# B&R Automation Studio project lab2_2
Automation Studio 4.5.2.102; technology packages: Acp10Arnc0 5.2.1

## Configuration Config1

CPU 4PP065.0571-P74, AutomationRuntime D4.52, Build 4.1.2, Vc V4.52.0, Safety 1.6

### Task classes (Cpu.sw)
```
Cyclic#1:
  ncsdcctrl <- ncsdcctrl.prg
Cyclic#2:
  Program <- Program.prg
DataObjects: Arnc0sys, Acp10sys
NcDataObjects: acp10etxen <- acp10etxen.dob, gmcipvar <- GmcIpUserConfig.gmcipvar.dob, gmcipfun <- GmcIpUserConfig.gmcipfun.dob, gmcipfub <- GmcIpUserConfig.gmcipfub.dob, gmcipubr <- GmcIpUserConfig.gmcipubr.dob, gmcipusm <- GmcIpUserConfig.gmcipusm.dob, gmcipui <- GmcIpUserConfig.gmcipui.dob, gmcipus <- GmcIpUserConfig.gmcipus.dob, gmcipuc <- GmcIpUserConfig.gmcipuc.dob, gmcipsys <- GmcIpConfig.gmcipsys.dob, gmciplbr <- GmcIpConfig.gmciplbr.dob, gmcipcbr <- GmcIpConfig.gmcipcbr.dob, gmciplsm <- GmcIpConfig.gmciplsm.dob, gmcipcsm <- GmcIpConfig.gmcipcsm.dob, gmcipcfg <- GmcIpConfig.gmcipcfg.dob, gmcipiec <- GmcIpConfig.gmcipiec.dob, gmciplog <- GmcIpConfig.gmciplog.dob, gmcipesm <- GmcIpConfig.gmcipesm.dob, gmcipmxd <- GmcIpConfig.gmcipmxd.dob, gmcipmx <- GmcIpConfig.gmcipmx.dob, gAxis01a <- gAxis01obj.gAxis01a.dob, gAxis01i <- gAxis01obj.gAxis01i.dob
Binaries: udbdef, TCData, iomap, asfw, Role, ashwac, sysconf, ashwd, User, arconfig, Arnc0map, acp10cfg, Acp10map, arnc0cfg
Libraries: Acp10man, Acp10par, NcGlobal, Acp10sdc, AsBrStr, Arnc0man, DataObj, AsArLog, sys_lib, FileIO, AsArProf, AsMem, brsystem, runtime, astime, Acp10_MC, Library, asieccon, powerlnk
```

### IoMap.iom - 4PP065_0571_P74/IoMap.iom
```iecst
VAR_CONFIG
	Cyclic#1.gAxis01_DrvIf.iLifeCnt AT %IB."X20SM1436a".LifeCnt;
	Cyclic#1.gAxis01_DrvIf.iDrvOK AT %IX."X20SM1436a".DrvOk01;
	Cyclic#1.gAxis01_DrvIf.oBoostCurrent AT %QX."X20SM1436a".BoostCurrent01;
	Cyclic#1.gAxis01_DrvIf.oStandStillCurrent AT %QX."X20SM1436a".StandstillCurrent01;
	Cyclic#1.gAxis01_DrvIf.oSetTime AT %QW."X20SM1436a".SetTime01;
	Cyclic#1.gAxis01_MotorStep0 AT %QW."X20SM1436a".Motor1Step0;
	Cyclic#1.gAxis01_DiDoIf.iLifeCntDriveEnable AT %IB."X20SM1436a".LifeCnt;
	Cyclic#1.gAxis01_DiDoIf.iLifeCntDriveReady AT %IB."X20SM1436a".LifeCnt;
	Cyclic#1.gAxis01_DiDoIf.iDriveReady AT %IX."X20SM1436a".DrvOk01;
	Cyclic#1.gAxis01_DiDoIf.oDriveEnable AT %QX."X20SM1436a".DriveEnable01;
	Cyclic#1.gAxis01_EncIf1.iLifeCnt AT %IB."X20SM1436a".LifeCnt;
	Cyclic#1.gAxis01_EncIf1.iEncOK AT %IX."X20SM1436a".EncOk01;
	Cyclic#1.gAxis01_EncIf1.iActPos AT %IW."X20SM1436a".ActPos01;
	Cyclic#1.gAxis01_EncIf1.iRefPulsePos AT %IW."X20SM1436a".RefPulsePos01;
	Cyclic#1.gAxis01_EncIf1.iRefPulseCnt AT %IB."X20SM1436a".RefPulseCnt01;
	Cyclic#1.gAxis01_EncIf1.iActTime AT %IW."X20SM1436a".ActTime01;
	::stateMachine.state AT %IW."8I64xxxxxxx.00x-1".ETAD_Input;
	::stateMachine.command AT %QW."8I64xxxxxxx.00x-1".CMDD_Output;
	::stateMachine.speed AT %QW."8I64xxxxxxx.00x-1".LFRD_Output;
	::doorSM.direction AT %IX."X20DI9371".DigitalInput01;
	::doorSM.sw1 AT %IX."X20DI9371".DigitalInput02;
	::doorSM.sw2 AT %IX."X20DI9371".DigitalInput03;
	::doorSM.sw3 AT %IX."X20DI9371".DigitalInput04;
	::doorSM.sw4 AT %IX."X20DI9371".DigitalInput05;
	::ledSM.led1 AT %QX."X20DO9322".DigitalOutput02;
	::ledSM.led2 AT %QX."X20DO9322".DigitalOutput03;
	::ledSM.led3 AT %QX."X20DO9322".DigitalOutput04;
	::ledSM.led4 AT %QX."X20DO9322".DigitalOutput05;
END_VAR
```

### Acp10cfg.ncc - 4PP065_0571_P74/Motion/Acp10cfg.ncc
```
NcConfiguration (Version=5.02.1, NcSwId=Acp10)
  ACP10CF1_typ:
    cnt_nettrc_rec_drive = 1500
    bufsize_trace_upload = 1200
    tc_nc_man_task = Cyclic #1
    glob_pv_as_ncobject = Yes
    ncsys_dl_broadcast = Yes
    ncsys_dl_acp_reset = Yes
    safemc_log_err_to_ax = Yes
    network_init:
      ncsw_init_execute = Yes
      automatic_execute = No
      node_nr_warning = Yes
      net_err_before_ncact = Yes
    nettrc:
      enter_parsecrec = Yes
      enter_ncaction = Yes
      save_ring_startidx = Yes
    cam_prof_download:
      cam_dat_dl_parallel = No
      tc_cam_dl_parallel = Task class for NC Manager task
    sdc_if[0]:
      if_name = SDC_IF1
      mc_broadcast_size = 800
      mc_broadcast_extdat = No
```

### Acp10map.ncm - 4PP065_0571_P74/Motion/Acp10map.ncm
```
NcMapping (NcSwId=Acp10)
  NcObject X20SM1436_ncAXIS1 (ModuleId=X20SM1436, ModuleAddress=SDC_IF1.ST1, Type=ncAXIS, Channel=1, AcoposSimulation=Off, Disabled=TRUE, ModuleDisabled=FALSE)
  NcObject gAxis01 (ModuleId=X20SM1436a, ModuleAddress=SDC_IF1.ST2, Type=ncAXIS, Channel=1, AcoposSimulation=Off, InitParameter=gAxis01i, AcoposParameter=gAxis01a, AdditionalData=CNC_Enabled="1" , Disabled=FALSE, ModuleDisabled=FALSE)
```

### Arnc0cfg.ncc - 4PP065_0571_P74/Motion/Arnc0cfg.ncc
```
NcConfiguration (Version=5.02.1, NcSwId=Arnc0)
  ARNC0CFG_typ:
    sampling_rate = 4000
    cnt_nettrc_rec_drive = 150
    bufsize_sys_trace = 16#00005000
    enable_mp_log = Yes
    tc_nc_man_task = Cyclic #1
    bg_load = 1
    glob_pv_as_ncobject = Yes
```

### Arnc0map.ncm - 4PP065_0571_P74/Motion/Arnc0map.ncm
```
NcMapping (NcSwId=Arnc0)
  NcObject CNC1 (Type=ncCNCSYS, Channel=1, AcoposSimulation=Off, Disabled=TRUE, ModuleDisabled=FALSE)
  NcObject CNC2 (Type=ncCNCSYS, Channel=2, AcoposSimulation=Off, Disabled=TRUE, ModuleDisabled=FALSE)
  NcObject CNC3 (Type=ncCNCSYS, Channel=3, AcoposSimulation=Off, Disabled=TRUE, ModuleDisabled=FALSE)
  NcObject CNC4 (Type=ncCNCSYS, Channel=4, AcoposSimulation=Off, Disabled=TRUE, ModuleDisabled=FALSE)
  NcObject CNC5 (Type=ncCNCSYS, Channel=5, AcoposSimulation=Off, Disabled=TRUE, ModuleDisabled=FALSE)
  NcObject CNC6 (Type=ncCNCSYS, Channel=6, AcoposSimulation=Off, Disabled=TRUE, ModuleDisabled=FALSE)
  NcObject CNC7 (Type=ncCNCSYS, Channel=7, AcoposSimulation=Off, Disabled=TRUE, ModuleDisabled=FALSE)
  NcObject CNC8 (Type=ncCNCSYS, Channel=8, AcoposSimulation=Off, Disabled=TRUE, ModuleDisabled=FALSE)
  NcObject CNC9 (Type=ncCNCSYS, Channel=9, AcoposSimulation=Off, Disabled=TRUE, ModuleDisabled=FALSE)
  NcObject CNC10 (Type=ncCNCSYS, Channel=10, AcoposSimulation=Off, Disabled=TRUE, ModuleDisabled=FALSE)
  NcObject CNC11 (Type=ncCNCSYS, Channel=11, AcoposSimulation=Off, Disabled=TRUE, ModuleDisabled=FALSE)
  NcObject CNC12 (Type=ncCNCSYS, Channel=12, AcoposSimulation=Off, Disabled=TRUE, ModuleDisabled=FALSE)
  NcObject CNC13 (Type=ncCNCSYS, Channel=13, AcoposSimulation=Off, Disabled=TRUE, ModuleDisabled=FALSE)
  NcObject CNC14 (Type=ncCNCSYS, Channel=14, AcoposSimulation=Off, Disabled=TRUE, ModuleDisabled=FALSE)
  NcObject CNC15 (Type=ncCNCSYS, Channel=15, AcoposSimulation=Off, Disabled=TRUE, ModuleDisabled=FALSE)
  NcObject CNC16 (Type=ncCNCSYS, Channel=16, AcoposSimulation=Off, Disabled=TRUE, ModuleDisabled=FALSE)
  NcObject CNC17 (Type=ncCNCSYS, Channel=17, AcoposSimulation=Off, Disabled=TRUE, ModuleDisabled=FALSE)
  NcObject CNC18 (Type=ncCNCSYS, Channel=18, AcoposSimulation=Off, Disabled=TRUE, ModuleDisabled=FALSE)
  NcObject CNC19 (Type=ncCNCSYS, Channel=19, AcoposSimulation=Off, Disabled=TRUE, ModuleDisabled=FALSE)
  NcObject CNC20 (Type=ncCNCSYS, Channel=20, AcoposSimulation=Off, Disabled=TRUE, ModuleDisabled=FALSE)
  NcObject CNC21 (Type=ncCNCSYS, Channel=21, AcoposSimulation=Off, Disabled=TRUE, ModuleDisabled=FALSE)
  NcObject CNC22 (Type=ncCNCSYS, Channel=22, AcoposSimulation=Off, Disabled=TRUE, ModuleDisabled=FALSE)
  NcObject CNC23 (Type=ncCNCSYS, Channel=23, AcoposSimulation=Off, Disabled=TRUE, ModuleDisabled=FALSE)
  NcObject CNC24 (Type=ncCNCSYS, Channel=24, AcoposSimulation=Off, Disabled=TRUE, ModuleDisabled=FALSE)
```

- Physical/Config1/4PP065_0571_P74/PvMap.vvm: same as Physical/Config1/4PP065_0571_P74/Cpu.per
## Logical view

Binary libraries used (declarations not repeated): operator, runtime, astime, AsIecCon, Acp10man 5.02.1, Acp10par 5.02.1, NcGlobal 5.02.1, Acp10sdc 5.02.1, AsBrStr, Arnc0man 5.02.1, DataObj, AsArLog, sys_lib, FileIO, AsArProf, AsMem, brsystem, Acp10_MC 5.02.1

### Global.var - Global variables
```iecst
VAR
	doorSM : DoorStateMachine;
	gAxis01 : ACP10AXIS_typ;
	gAxis01_DiDoIf : SdcDiDoIf_typ := (0);
	gAxis01_DrvIf : SdcDrvIf16_typ := (0);
	gAxis01_EncIf1 : SdcEncIf16_typ := (0);
	gAxis01_HW : SdcHwCfg_typ := (0);
	gAxis01_MotorStep0 : INT := (0);
	ledSM : LedStateMachine;
	stateMachine : DriveStateMachine;
END_VAR
```


### Data object Logical/acp10etxen (Ett)

- acp10etxen.ett (not shown)

### Program Logical/ncsdcctrl (IEC)

#### ncsdcctrlCyclic.st
```iecst
PROGRAM _CYCLIC

(* ### BEGIN gAxis01 ### *)

(* life counter emulation of digital inputs *)
      gAxis01_DiDoIf.iLifeCntReference := gAxis01_DiDoIf.iLifeCntReference + 1;
      gAxis01_DiDoIf.iLifeCntNegHwEnd  := gAxis01_DiDoIf.iLifeCntNegHwEnd  + 1;
      gAxis01_DiDoIf.iLifeCntPosHwEnd  := gAxis01_DiDoIf.iLifeCntPosHwEnd  + 1;

(* default function model of ACOPOSmicro: convert absolute steps to delta steps - overflow save delta calculation *)
      gAxis01_MotorStep0 := gAxis01_DrvIf.oSetPos - gAxis01_oSetPosOld;
      gAxis01_oSetPosOld := gAxis01_DrvIf.oSetPos;

(* ### END gAxis01 ### *)

END_PROGRAM
```

#### ncsdcctrlInit.st
```iecst
PROGRAM _INIT

(* ### BEGIN gAxis01 ### *)

(* initialize general interfaces *)
      gAxis01.size := gAxis01.size;
      gAxis01_HW.DrvIf_Typ := ncSDC_DRVSM16;
      brsstrcpy( ADR(gAxis01_HW.DrvIf_Name[0]), ADR('gAxis01_DrvIf') );
      gAxis01_HW.DiDoIf_Typ := ncSDC_DIDO;
      brsstrcpy( ADR(gAxis01_HW.DiDoIf_Name[0]), ADR('gAxis01_DiDoIf') );
      gAxis01_HW.EncIf1_Typ := ncSDC_ENC16;
      brsstrcpy( ADR(gAxis01_HW.EncIf1_Name[0]), ADR('gAxis01_EncIf1') );
      gAxis01_EncIf1.iLifeCnt := gAxis01_EncIf1.iLifeCnt;

(* initialize old-value for delta step calculation *)
      gAxis01_oSetPosOld := gAxis01_DrvIf.oSetPos;

(* ### END gAxis01 ### *)

END_PROGRAM
```

#### ncsdcctrl.var
```iecst
VAR
	gAxis01_oSetPosOld : INT := 0;
END_VAR
```

### Data object Logical/GmcIpConfig/gmcipsys (Cnc, version 5.02.1)

#### gmcipsys.cnc
```
LANGS (defaultLangId=1, defaultDataLangId=3)
  CMDQUEUE (BufferSize=15)
  MEM (ReserveMB=5, LimitPercent=80%)
  EXEC (InstrBurstBG=200, CycleBurstBG=0, Stack=16384, MinorStack=2048, EStack=1024)
  LOAD (ReadLineBurstMax=100, ReadLineBurstMin=20, ParseLineBurstMax=10, ParseLineBurstMin=2, RuntimeIOBlocking=No)
  DISABLE_MSG = 15238 
    15336 
    15337 
    15666 
    15784 
    15864 
    15740
  LANG (langId=1, langName=B&R GCode, langModule=ailgcode)
    LANGCONFIG gmciplbr
    LANGCONFIG gmcipcbr
    LANGCONFIG gmcipubr
    FILEEXT .cnc
    FILEEXT .prg
    MAINSEARCHPATH $ (FileDevice=CNC_PrgDir)
    MAINSEARCHPATH $ (DataObject=Yes)
    INCLUDEPATH $ (FileDevice=CNC_PrgDir)
    INCLUDEPATH $ (DataObject=Yes)
  LANG (langId=2, langName=Alternative Language 1 GCode, langModule=ailgcode)
    LANGCONFIG gmciplsm
    LANGCONFIG gmcipcbr
    LANGCONFIG gmcipcsm
    LANGCONFIG gmcipusm
    FILEPREFIX = _N_
    FILEEXT = .MPF
    FILEEXT = _MPF
    FILEEXT = .SPF
    FILEEXT = _SPF
    MAINSEARCHPATH = \$ (FileDevice=CNC_PrgDir)
    MAINSEARCHPATH = \_N_MPF_DIR\$ (FileDevice=CNC_PrgDir)
    MAINSEARCHPATH = \_N_SPF_DIR\$ (FileDevice=CNC_PrgDir)
    MAINSEARCHPATH = $ (DataObject=1)
    INCLUDEPATH = \$ (FileDevice=CNC_PrgDir)
    INCLUDEPATH = \_N_SPF_DIR\$ (FileDevice=CNC_PrgDir)
    INCLUDEPATH = \_N_MPF_DIR\$ (FileDevice=CNC_PrgDir)
    INCLUDEPATH = $ (DataObject=1)
  LANG (langId=3, langName=IEC-ST, langModule=ailgcode)
    LANGCONFIG gmcipiec
    LANGCONFIG gmcipmx (RequireFnIgnore=MXConvertOrient)
    LANGCONFIG gmcipui (IfNotExist=Warn)
    FILEEXT .typ (DeclScope=IP_GLOBAL)
    FILEEXT .var (DeclScope=IP_GLOBAL)
    FILEEXT .fun (DeclScope=IP_GLOBAL)
    FILEEXT .iec (DeclScope=IP_LOCAL)
    FILEEXT .st (DeclScope=IP_LOCAL)
    FILEEXT _iec (DeclScope=IP_LOCAL)
    MAINSEARCHPATH = \$ (FileDevice=IEC_PrgDir)
    MAINSEARCHPATH = \$ (FileDevice=CNC_PrgDir)
    MAINSEARCHPATH \TYP\$ (FileDevice=CNC_PrgDir, DataObject=No)
    INCLUDEPATH = \$ (FileDevice=IEC_PrgDir)
    INCLUDEPATH = \$ (FileDevice=CNC_PrgDir)
    INCLUDEPATH \TYP\$ (FileDevice=CNC_PrgDir, DataObject=No)
  XML_INCLUDE gmcipus (IfNotExist=Warn)
```

### Data object Logical/GmcIpConfig/gmciplbr (Cnc, version 5.02.1)

#### gmciplbr.cnc
```
Root (LangModule=ailgcode, Version=1.0)
  BuiltInProcs:
    cancel = beginpathsynch
        StopCyclicGroups(:${*}:);
      endpathsynch (MinArgs=1, MaxArgs=*)
  BuiltInFns (PatternSuffix=:\[)
    ABS = Abs(:$[1]:) (NumArgs=1, Inline=Yes)
    SQR = ($[1] * $[1]) (NumArgs=1)
    ACOS = ACos(:$[1]:) (NumArgs=1, Inline=Yes)
    ASIN = ASin(:$[1]:) (NumArgs=1, Inline=Yes)
    ATAN = ATan(:$[1]:) (NumArgs=1, Inline=Yes)
    COS = Cos(:$[1]:) (NumArgs=1, Inline=Yes)
    DEXP = DExp(:$[1]:) (NumArgs=1, Inline=Yes)
    EXP = Exp(:$[1]:) (NumArgs=1, Inline=Yes)
    FIX = Fix(:$[1]:) (NumArgs=1, Inline=Yes)
    FRACT = Fract(:$[1]:) (NumArgs=1, Inline=Yes)
    FUP = Fup(:$[1]:) (NumArgs=1, Inline=Yes)
    INV = ~($[1]) (NumArgs=1, Inline=Yes)
    LN = Ln(:$[1]:) (NumArgs=1, Inline=Yes)
    LOG = Log(:$[1]:) (NumArgs=1, Inline=Yes)
    ROUND = ToInt(:$[1]:) (NumArgs=1, Inline=Yes)
    SIN = Sin(:$[1]:) (NumArgs=1, Inline=Yes)
    SQRT = Sqrt(:$[1]:) (NumArgs=1, Inline=Yes)
    TAN = Tan(:$[1]:) (NumArgs=1, Inline=Yes)
    BOOL = ToBool(:$[1]:) (NumArgs=1, Inline=Yes)
    INT = Fix(:$[1]:) (NumArgs=1, Inline=Yes)
    ADR = Adr(:\$[1]:) (NumArgs=1, Inline=Yes)
    SIZEOF = Sizeof(:\$[1]:) (NumArgs=1, Inline=Yes)
    NUM_LOADED_FILES = NumLoadedFiles(::) (NumArgs=0)
    NUM_LOADED_PROG_FILES = NumLoadedProgFiles(::) (NumArgs=0)
    MEM_SIZE_IP_ALL = MemSizeIpInstAll(::) (NumArgs=0)
    MEM_SIZE_IP_LIB = MemSizeIpInst(::) (NumArgs=0)
    MEM_SIZE_SHLIB = MemSizeShLib(::) (NumArgs=0)
    MEM_SIZE_FILE = MemSizeFile(:$[1]:) (MinArgs=0, MaxArgs=1)
    MEM_SIZE_IP_STACK_SPACE = MemStackSpace(::) (NumArgs=0)
  AxesSpec:
    AxisRef = $\s*=\s*AC (Mode=3)
    AxisRef = $\s*=\s*IC (Mode=4)
  PVMacros:
    RDISABLE (ArrayDims=0, Group=500)
      CALL = @#job->sa.keep_alive = 1;
        @#thread.sa_keep_alive = 1; (Inline=Yes)
  Parameters:
    R (IndexType=RParamIndex, ValueType=FLOAT)
      ARG (ref=EXPR, DataType=RParamIndex)
    P (IndexType=RParamIndex, ValueType=FLOAT)
      ARG (ref=EXPR, DataType=RParamIndex)
    EXB (IndexType=EXParamIndex, ValueType=Byte)
      ARG (ref=EXPR, DataType=EXParamIndex)
    EXW (IndexType=EXParamIndex, ValueType=Word)
      ARG (ref=EXPR, DataType=EXParamIndex)
    EXL (IndexType=EXParamIndex, ValueType=Long)
      ARG (ref=EXPR, DataType=EXParamIndex)
    EXF (IndexType=EXFParamIndex, ValueType=FLOAT)
      ARG (ref=EXPR, DataType=EXFParamIndex)
    MW (Synchronous=Yes, IndexType=MParamIndex, ValueType=Word)
      ARG (ref=EXPR, DataType=MParamIndex)
    ML (Synchronous=Yes, IndexType=MParamIndex, ValueType=Long)
      ARG (ref=EXPR, DataType=MParamIndex)
    MF (Synchronous=Yes, IndexType=MParamIndex, ValueType=FLOAT)
      ARG (ref=EXPR, DataType=MParamIndex)
  PrimTypes (PatternSuffix=:[^\[], MapIECTypes=Yes)
  Preprocess:
    PP_RULE_FRAME_I (Search=$FRAME_I, Replace=[1,0,0,0,1,0,0,0,1,0,0,0])
    PP_RULE_FRAME_DEF (IsPattern=Yes, Search=FRAME:[^\w\d], Replace=LREAL{12})
  FubTemplates:
    StdFubTemplate (IsDefault=Yes, Inline=Yes)
      Arg (ref=FUBINST, DataType=FLOAT)
      Arg (ref=FUBERRLEV, DataType=FLOAT)
      Arg (ref=PATHSYNCH, DataType=FLOAT)
      Arg (ref=BLOCKING, DataType=FLOAT)
  SynchActions:
    SABlocks:
      default (IsDefault=Yes)
        cyclic (Inline=Yes)
          Arg (ref=ACTIONS, DataType=STATEMENTS)
          Arg (ref=ID, DataType=FLOAT, DefaultInt=-1, MinCount=0, MaxCount=1)
      whenever:
        cyclic (Inline=Yes)
          Arg (ref=COND, DataType=FLOAT)
          Arg (ref=ACTIONS, DataType=STATEMENTS)
          Arg (ref=ID, DataType=FLOAT, DefaultInt=-1, MinCount=0, MaxCount=1)
      when:
        cyclic (Inline=Yes)
          Arg (ref=COND, DataType=FLOAT)
          Arg (ref=ACTIONS, DataType=STATEMENTS)
          Arg (ref=ID, DataType=FLOAT, DefaultInt=-1, MinCount=0, MaxCount=1)
      every:
        cyclic (Inline=Yes)
          Arg (ref=COND, DataType=FLOAT)
          Arg (ref=ACTIONS, DataType=STATEMENTS)
          Arg (ref=ID, DataType=FLOAT, DefaultInt=-1, MinCount=0, MaxCount=1)
      from:
        cyclic (Inline=Yes)
          Arg (ref=COND, DataType=FLOAT)
          Arg (ref=ACTIONS, DataType=STATEMENTS)
          Arg (ref=ID, DataType=FLOAT, DefaultInt=-1, MinCount=0, MaxCount=1)
    NonModalActivation:
      Start = @#thread.sa_last_keep_alive = 1;
        ActivateCyclicGroup(:-1:);
      Stop = WaitStopCyclicGroups(:(:-1:):);
  ParserData (NestedComments=Yes, DefaultCaseSensitive=No, CommentsSpanLines=No, SubDeclsLocalToFile=Yes, ProgDeclsLocalToFile=Yes, AllowUnprefixedFileCalls=No, LocalVarScopeForMainProg=No, FileScopeVarsVisibleInSub=Yes, MainPrgReturnAtNextMainPrgHdr=Yes, MaxSizePassByValue=1024, AllowVarReadBeforeAssign=No, AllowArrayRefWithoutIndex=Yes, AllowStructMemberAutoDereference=Yes, AllowVariableAutoDereference=Yes, AllowIgnoredExtraSubArgs=Yes, EnableStringCharacterIndexing=Yes, OnMacroRedefinition=Warn, CheckFileTimestampBeforeCalls=Yes)
    TKG_END_OF_LINE = \n (IsPattern=No)
    TKG_LINE_CONTINUE = \ (IsPattern=No, FileXLInvalid=Yes)
    TKG_LINE_BREAK = @@
    TKG_ARITH_BINARY_MODULO = MOD
    TKG_TRUE = TRUE:\W (IsPattern=Yes)
    TKG_FALSE = FALSE:\W (IsPattern=Yes)
    TKG_PAREVAL_MODAL_ID = ID:[\s=] (FileXLInvalid=Yes, IsPattern=Yes)
    TKG_OPEN_COMMENT = (
    TKG_CLOSE_COMMENT = )
    TKG_OPEN_BRACKET = [
    TKG_COMMA = ,
    TKG_CLOSE_BRACKET = ]
    TKG_OPEN_INDEXBRACKET = {
    TKG_CLOSE_INDEXBRACKET = }
    TKG_NUMBER = \d+\.\d+|\d+\.:[^\.] (IsPattern=Yes)
    TKG_INTEGER = \d+ (IsPattern=Yes)
    TKG_FRACTION = \.\d+ (IsPattern=Yes)
    TKG_DOT = \.:\w (IsPattern=Yes, FollowedBy=TKG_STRUCT_MEMBER_REF)
    TKG_STRUCT_MEMBER_REF = \w|\w[\w\d]+ (IsPattern=Yes, Restricted=Yes)
    TKG_NUMBER_EXP = EX:[\s\d\+\-\.] (IsPattern=Yes)
    TKG_MACRO_DEFINE_GLOBAL = define\s+ip_global:\s (IsPattern=Yes, FollowedBy=TKG_MACRO_NAME)
    TKG_MACRO_DEFINE = define\s+local:\s|define:\s (IsPattern=Yes, FollowedBy=TKG_MACRO_NAME)
    TKG_MACRO_UNDEFINE = undefine:\s (IsPattern=Yes, FollowedBy=TKG_MACRO_NAME)
    TKG_MACRO_AS = as:[\s\n] (IsPattern=Yes, FollowedBy=TKG_MACRO_TEXT)
    TKG_MACRO_NAME = [$\w][$\w\d]+ (Restricted=Yes, IsPattern=Yes)
    TKG_MACRO_TEXT = . (Restricted=Yes, IsPattern=Yes)
    TKG_BUILTIN_NUM_FN_NAME
    _TKG_LABEL_DEF1:
      TKG_LABEL_DEF = L[\w\d]+:\:[^\w\d] (IsPattern=Yes, FollowedBy=TKG_LABEL_SUFFIX)
    TKG_SUBPROG_START = %:L (FileXLInvalid=Yes, IsPattern=Yes, FollowedBy=TKG_SUBPROG_NAME)
    TKG_SUBPROG_NAME = L\d+ (IsPattern=Yes, Restricted=Yes)
    TKG_SUBPROG_CALL = L:L\d (IsPattern=Yes, FollowedBy=TKG_SUBPROG_NAME)
    TKG_SUBPROG_PROTO = %D:L (IsPattern=Yes, FollowedBy=TKG_SUBPROG_NAME)
    TKG_SUBCALL_REPEAT_PREFIX = O:[\s\d] (IsPattern=Yes, FollowedBy=TKG_INTEGER)
    TKG_EXTERN = EXTERN:\s (IsPattern=Yes, FollowedBy=TKG_PROG_FILE_NAME)
    TKG_ARG_PASSBYREF = VAR\s (IsPattern=Yes)
    TKG_SET_MODAL_SUB = MCALL:\W (FileXLInvalid=Yes, IsPattern=Yes)
    TKG_PROG_START = %:\d (IsPattern=Yes, FollowedBy=TKG_PROG_NAME)
    TKG_PROG_NAME = \d+ (IsPattern=Yes, Restricted=Yes)
    TKG_PROG_CALL = L:[^L] (IsPattern=Yes, FollowedBy=TKG_PROG_FILE_NAME)
    TKG_PROG_FILE_NAME = [\^#&@']?[\w\d\.\\]+:[^\w\d\.\\\:]|[\^#][\w\d]+\:[\w\d\.\\]+ (IsPattern=Yes, Restricted=Yes)
    TKG_SUPPRESS_SINGLE_STEP = NOHALT
    TKG_NC_BLOCK_PREFIX = N:[\d\s] (IsPattern=Yes)
    TKG_PARAM_PREFIX = R:\d|P:\d|M[WLF]:\d|EX[WLBF]:\d (IsPattern=Yes)
    TKG_SUBRANGE = ..
    TKG_G_CODE_PREFIX = G:[\s\d] (IsPattern=Yes)
    TKG_M_CODE_PREFIX = M:[\s\d\[] (IsPattern=Yes)
    TKG_PAREVAL_DO = do:\s (FileXLInvalid=Yes, IsPattern=Yes)
    TKG_GOTO = $GOTO:\s (FileXLInvalid=Yes, IsPattern=Yes, OptFollowedBy=TKG_GOTO_DEST)
    TKG_GOTO_DEST = \w[\w\d]* (IsPattern=Yes, Restricted=Yes)
    TKG_LOGICAL_BINARY_AND = &&
    TKG_LOGICAL_BINARY_OR = ||
    TKG_LOGICAL_BINARY_XOR = XOR
    TKG_STRING_CONCAT = <<
    TKG_COMP_BINARY_GREATER_THAN_OR_EQ = >=
    TKG_COMP_BINARY_LESS_THAN_OR_EQ = <=
    TKG_COMP_BINARY_EQUAL_TO = ==
    TKG_COMP_BINARY_NOT_EQUAL_TO = !=
    TKG_COMP_BINARY_GREATER_THAN = >
    TKG_COMP_BINARY_LESS_THAN = <
    TKG_ASSIGN_EQ = =
    TKG_LOGICAL_UNARY_NOT = !
    TKG_BITWISE_BINARY_AND = &
    TKG_BITWISE_BINARY_OR = |
    TKG_BITWISE_BINARY_XOR = ^
    TKG_BITWISE_UNARY_COMPLEMENT = ~
    TKG_ARITH_BINARY_PLUS = +
    TKG_ARITH_BINARY_MINUS = -
    TKG_ARITH_BINARY_POWER = **
    TKG_ARITH_BINARY_MULTIPLY = *
    TKG_ARITH_BINARY_DIVIDE = /
    TKG_PATHSYNCH_REC_IEC = $DO_PATH_SYNCH (FileXLInvalid=Yes)
    TKG_PATHSYNCH_END = $END_PATH_SYNCH (FileXLInvalid=Yes)
    TKG_PATHSYNCH_IPEVAL = $IP_EVAL (FileXLInvalid=Yes)
    TKG_IF = $IF (FileXLInvalid=Yes)
    TKG_THEN = $THEN (FileXLInvalid=Yes)
    TKG_BLOCK_ELSEIF = $ELSEIF (FileXLInvalid=Yes)
    TKG_BLOCK_ELSE = $ELSE (FileXLInvalid=Yes)
    TKG_BLOCK_ENDIF = $ENDIF (FileXLInvalid=Yes)
    TKG_SWITCH = $SWITCH (FileXLInvalid=Yes)
    TKG_SWITCH_CASE = $CASE (FileXLInvalid=Yes)
    TKG_SWITCH_DEFAULT = $DEFAULT (FileXLInvalid=Yes)
    TKG_ENDSWITCH = $ENDSWITCH (FileXLInvalid=Yes)
    TKG_FOR = $FOR (FileXLInvalid=Yes)
    TKG_ENDFOR = $ENDFOR (FileXLInvalid=Yes)
    TKG_WHILE = $WHILE (FileXLInvalid=Yes)
    TKG_ENDWHILE = $ENDWHILE (FileXLInvalid=Yes)
    TKG_DO = $DO (FileXLInvalid=Yes)
    TKG_ENDDO = $ENDDO (FileXLInvalid=Yes)
    TKG_BREAK = $BREAK (FileXLInvalid=Yes)
    TKG_CONTINUE = $CONTINUE (FileXLInvalid=Yes)
    TKG_PRIM_TYPE (IsPattern=Yes)
    TKG_PV_DECL = def:\s (IsPattern=Yes)
    TKG_PV_UNDECL = ~def:\s (IsPattern=Yes)
    TKG_PV_DECL_REF = \w[\w\d\.\:\*]+|\w (IsPattern=Yes, Restricted=Yes)
    TKG_VARSCOPE_IP_LOCAL = local:[\s\n] (IsPattern=Yes)
    TKG_VARSCOPE_IP_GLOBAL = ip_global:[\s\n] (IsPattern=Yes)
    TKG_VARSCOPE_NC_GLOBAL = nc_global:[\s\n] (IsPattern=Yes)
    TKG_VARSCOPE_PLC_GLOBAL = plc_global:[\s\n] (IsPattern=Yes)
    TKG_VAR_RETAIN = retain:\s (IsPattern=Yes)
    TKG_VARSYNCH_IP = ip_synch:\s (IsPattern=Yes)
    TKG_VARSYNCH_PATH = path_synch:\s (IsPattern=Yes)
    TKG_LABEL_DEF = \w:\:|\w[\w\d]+:\: (IsPattern=Yes, FollowedBy=TKG_LABEL_SUFFIX)
    TKG_LABEL_SUFFIX = : (Restricted=Yes)
    TKG_FUB_DECL = fub:\s (IsPattern=Yes)
    TKG_FUB_ERR_LEV_1 = error_level_1:\s (IsPattern=Yes)
    TKG_FUB_ERR_LEV_2 = error_level_2:\s (IsPattern=Yes)
    TKG_FUB_ERR_LEV_3 = error_level_3:\s (IsPattern=Yes)
    TKG_FUB_ERR_LEV_4 = error_level_4:\s (IsPattern=Yes)
    TKG_FUB_BLOCKING = blocking:\s (IsPattern=Yes)
    TKG_FUB_NON_BLOCKING = non_blocking:\s (IsPattern=Yes)
    TKG_IEC_TYPED_VALUE = #[\w\d]+ (IsPattern=Yes)
    TKG_REFERENCE = ref:[\s\n]|reference:[\s\n] (IsPattern=Yes, FollowedBy=TKG_IEC_TO)
    TKG_IEC_TO = to:[\s\n] (IsPattern=Yes, Restricted=Yes)
    TKG_ACCESS = ACCESS:[\s\n] (IsPattern=Yes)
    TKG_WORD = \w|\w[\w\d\.]+ (IsPattern=Yes)
  StringChars (AsciiStringStart=", UTF16StringStart=W", UTF16StringEnd=")
    EscapeSeq (Search=$N, ReplaceValue=10)
    EscapeSeq (Search=$L, ReplaceValue=10)
    EscapeSeq (Search=$P, ReplaceValue=12)
    EscapeSeq (Search=$R, ReplaceValue=13)
    EscapeSeq (Search=$T, ReplaceValue=9)
    EscapeSeq (Search=$Q, ReplaceStr=")
    EscapeSeq (Search=$', ReplaceStr=')
    EscapeSeq (Search=$", ReplaceStr=")
    EscapeSeq (Search=$[\dA-Fa-f]+, IsPattern=Yes, ReplaceEncodingBase=16)
    EscapeSeq (Search=$$, ReplaceStr=$)
    EscapeSeq (Search=$, ReplaceStr=)
```

### Data object Logical/GmcIpConfig/gmcipcbr (Cnc, version 5.02.1)

- gmcipcbr.cnc (not shown)

### Data object Logical/GmcIpConfig/gmciplsm (Cnc, version 5.02.1)

#### gmciplsm.cnc
```
Root (LangModule=ailgcode, Version=1.0)
  PrimTypes (CaseSensitive=No)
    REAL (BRType=LREAL)
    INT (BRType=DINT)
    CHAR (BRType=USINT)
    BOOL (BRType=BOOL)
    STRING (BRType=STRING)
    AXIS (BRType=AXIS)
    BR_LREAL (BRType=LREAL)
    BR_REAL (BRType=REAL)
    BR_UDINT (BRType=UDINT)
    BR_DINT (BRType=DINT)
    BR_UINT (BRType=UINT)
    BR_INT (BRType=INT)
    BR_USINT (BRType=USINT)
    BR_SINT (BRType=SINT)
    BR_BOOL (BRType=BOOL)
    BR_TIME (BRType=TIME)
    BR_DATE_AND_TIME (BRType=DATE_AND_TIME)
  Preprocess:
    PP_RULE_NCK (Search=NCK , Replace=nc_global )
    PP_RULE_CHAN (Search=CHAN , Replace=ip_global )
    PP_RULE_FRAME_I (Search=$FRAME_I, Replace=(1,0,0,0,1,0,0,0,1,0,0,0))
    PP_RULE_FRAME_DEF (IsPattern=Yes, Search=FRAME:[^\w\d], Replace=REAL[12])
  BuiltInProcs:
    cancel = beginpathsynch
        StopCyclicGroups(:${*}:);
      endpathsynch (MinArgs=1, MaxArgs=*)
    RET = #next_motion.Command = MPCMD_SET_M_FCT;
      #next_motion.Data.I4_value = 17;
      PushPacket(::);
      ReturnTo(:${*}:); (MinArgs=0, MaxArgs=4, Eval=Early, Inline=Yes)
  BuiltInFns:
    ABS = Abs(:$[1]:) (NumArgs=1, Inline=Yes)
    SIN = Sin(:$[1]:) (NumArgs=1, Inline=Yes)
    COS = Cos(:$[1]:) (NumArgs=1, Inline=Yes)
    TAN = Tan(:$[1]:) (NumArgs=1, Inline=Yes)
    ASIN = ASin(:$[1]:) (NumArgs=1, Inline=Yes)
    ACOS = ACos(:$[1]:) (NumArgs=1, Inline=Yes)
    ATAN = ATan(:$[1]:) (NumArgs=1, Inline=Yes)
    ATAN2 = ATan2(:$[1],$[2]:) (NumArgs=2, Inline=Yes)
    SQRT = Sqrt(:$[1]:) (NumArgs=1, Inline=Yes)
    POT = (($[1])*($[1])) (NumArgs=1, Inline=Yes)
    TRUNC = Fix(:$[1]:) (NumArgs=1, Inline=Yes)
    ROUND = Round(:$[1]:) (NumArgs=1, Inline=Yes)
    LN = Ln(:$[1]:) (NumArgs=1, Inline=Yes)
    EXP = Exp(:$[1]:) (NumArgs=1, Inline=Yes)
    MINVAL = MinVal(:$[1], $[2]:) (NumArgs=2, Inline=Yes)
    MAXVAL = MaxVal(:$[1], $[2]:) (NumArgs=2, Inline=Yes)
    BOUND = Bounds(:$[1], $[2], $[3]:) (NumArgs=3, Inline=Yes)
    TO_BOOL = ToBool(:$[1]:) (NumArgs=1, Inline=Yes)
    TO_INT = ToInt(:$[1]:) (NumArgs=1, Inline=Yes)
    TO_CHAR = ToChar(:$[1]:) (NumArgs=1, Inline=Yes)
    TO_REAL = ToLReal(:$[1]:) (NumArgs=1, Inline=Yes)
    TO_FLOAT = ToFloat(:$[1]:) (NumArgs=1, Inline=Yes)
    DEFINED = Defined(:$[1]:) (NumArgs=1, Inline=Yes)
    TIME_MS = TimeMs(::) (NumArgs=0)
    SET = ${*} (MinArgs=0, MaxArgs=*, Inline=Yes)
    REP = ArrayRep(:${*}:) (MinArgs=1, MaxArgs=2, Inline=Yes)
    ADR = Adr(:\$[1]:) (NumArgs=1, Inline=Yes)
    SIZEOF = Sizeof(:\$[1]:) (NumArgs=1, Inline=Yes)
    NUM_LOADED_FILES = NumLoadedFiles(::) (NumArgs=0)
    NUM_LOADED_PROG_FILES = NumLoadedProgFiles(::) (NumArgs=0)
    MEM_SIZE_IP_ALL = MemSizeIpInstAll(::) (NumArgs=0)
    MEM_SIZE_IP_LIB = MemSizeIpInst(::) (NumArgs=0)
    MEM_SIZE_SHLIB = MemSizeShLib(::) (NumArgs=0)
    MEM_SIZE_FILE = MemSizeFile(:$[1]:) (MinArgs=0, MaxArgs=1)
    MEM_SIZE_IP_STACK_SPACE = MemStackSpace(::) (NumArgs=0)
  AxesSpec:
    AxisRef = $\s*=\s*AC (Mode=3)
    AxisRef = $\s*=\s*IC (Mode=4)
  PVMacros:
    SBLOF (ArrayDims=0, Group=500)
      CALL = #call->forbid_stepping = 1; (Inline=Yes)
    SBLON (ArrayDims=0, Group=500)
      CALL = #call->forbid_stepping = 0; (Inline=Yes)
    DISPLOF (ArrayDims=0, Group=500)
      CALL = #call->forbid_display = 1; (Inline=Yes)
    DISPLON (ArrayDims=0, Group=500)
      CALL = #call->forbid_display = 0; (Inline=Yes)
    RDISABLE (ArrayDims=0, Group=500)
      CALL = @#job->sa.keep_alive = 1;
        @#thread.sa_keep_alive = 1; (Inline=Yes)
    P_SUBPAR $P_SUBPAR (ArrayDims=1, Group=500)
      GET = return ArgNumIsDefined(:$[1]:);
    P_STACK $P_STACK:
      GET = return UserCallDepth(::);
  FubTemplates:
    StdFubTemplate (IsDefault=Yes, Inline=Yes)
      Arg (ref=FUBINST, DataType=FLOAT)
      Arg (ref=FUBERRLEV, DataType=FLOAT)
      Arg (ref=PATHSYNCH, DataType=FLOAT)
      Arg (ref=BLOCKING, DataType=FLOAT)
  SynchActions:
    SABlocks:
      default (IsDefault=Yes)
        cyclic (Inline=Yes)
          Arg (ref=ACTIONS, DataType=STATEMENTS)
          Arg (ref=ID, DataType=FLOAT, DefaultInt=-1, MinCount=0, MaxCount=1)
      whenever:
        cyclic (Inline=Yes)
          Arg (ref=COND, DataType=FLOAT)
          Arg (ref=ACTIONS, DataType=STATEMENTS)
          Arg (ref=ID, DataType=FLOAT, DefaultInt=-1, MinCount=0, MaxCount=1)
      when:
        cyclic (Inline=Yes)
          Arg (ref=COND, DataType=FLOAT)
          Arg (ref=ACTIONS, DataType=STATEMENTS)
          Arg (ref=ID, DataType=FLOAT, DefaultInt=-1, MinCount=0, MaxCount=1)
      every:
        cyclic (Inline=Yes)
          Arg (ref=COND, DataType=FLOAT)
          Arg (ref=ACTIONS, DataType=STATEMENTS)
          Arg (ref=ID, DataType=FLOAT, DefaultInt=-1, MinCount=0, MaxCount=1)
      from:
        cyclic (Inline=Yes)
          Arg (ref=COND, DataType=FLOAT)
          Arg (ref=ACTIONS, DataType=STATEMENTS)
          Arg (ref=ID, DataType=FLOAT, DefaultInt=-1, MinCount=0, MaxCount=1)
    NonModalActivation:
      Start = @#thread.sa_last_keep_alive = 1;
        ActivateCyclicGroup(:-1:);
      Stop = WaitStopCyclicGroups(:(:-1:):);
  ParserData (NestedComments=Yes, DefaultCaseSensitive=No, CommentsSpanLines=No, SubDeclsLocalToFile=Yes, ProgDeclsLocalToFile=Yes, AllowUnprefixedFileCalls=Yes, AllowUnprefixedSubCalls=Yes, LocalVarScopeForMainProg=No, FileScopeVarsVisibleInSub=Yes, MainPrgReturnAtNextMainPrgHdr=Yes, AllowVarReadBeforeAssign=No, AllowArrayRefWithoutIndex=Yes, AllowNamedFnArgs=Yes, AllowBuiltinFnArgsOutOfSequence=Yes, AllowBuiltInProcCallWithoutBrackets=Yes, AllowBuiltInFnCallWithoutBrackets=No, AllowPLCFnCallWithoutBrackets=No, AllowStructMemberAutoDereference=Yes, AllowVariableAutoDereference=Yes, EnableStringCharacterIndexing=Yes, AllowIgnoredExtraSubArgs=Yes, OnMacroRedefinition=Error, CheckFileTimestampBeforeCalls=Yes)
    TKG_END_OF_LINE = \n (IsPattern=No)
    TKG_LINE_CONTINUE = \ (IsPattern=No, FileXLInvalid=Yes)
    TKG_LINE_BREAK = @@
    TKG_OPEN_COMMENT = ;
    TKG_CLOSE_COMMENT
    TKG_TRUE = TRUE:\W (IsPattern=Yes)
    TKG_FALSE = FALSE:\W (IsPattern=Yes)
    TKG_PAREVAL_MODAL_ID = ID:[\s=] (FileXLInvalid=Yes, IsPattern=Yes)
    TKG_MACRO_DEFINE_GLOBAL = define\s+ip_global:\s (IsPattern=Yes, FollowedBy=TKG_MACRO_NAME)
    TKG_MACRO_DEFINE = define\s+local:\s|define:\s (IsPattern=Yes, FollowedBy=TKG_MACRO_NAME)
    TKG_MACRO_UNDEFINE = undefine:\s (IsPattern=Yes, FollowedBy=TKG_MACRO_NAME)
    TKG_MACRO_AS = as:[\s\n] (IsPattern=Yes, FollowedBy=TKG_MACRO_TEXT)
    TKG_PROG_START = %:[^L] (IsPattern=Yes, CaseSensitive=Yes, FollowedBy=TKG_PROG_NAME)
    TKG_PROG_NAME = [\w\d]+ (IsPattern=Yes, Restricted=Yes)
    TKG_SET_MODAL_SUB = MCALL:\W (FileXLInvalid=Yes, IsPattern=Yes)
    TKG_INDIR_PROG_CALL = CALL:\s (IsPattern=Yes)
    TKG_INDIR_PROG_BLOCK = BLOCK:\s (FileXLInvalid=Yes, IsPattern=Yes)
    TKG_PROC_START = PROC:\s (FileXLInvalid=Yes, IsPattern=Yes, FollowedBy=TKG_PROC_NAME)
    TKG_PROC_NAME = \w[\w\d]+ (IsPattern=Yes, Restricted=Yes)
    TKG_ARG_PASSBYREF = VAR:\s (IsPattern=Yes)
    TKG_SUBPROG_PROTO = INTERN:\s (IsPattern=Yes, FollowedBy=TKG_SUBPROG_NAME)
    TKG_SUBPROG_START = SUB\s|%:L (FileXLInvalid=Yes, IsPattern=Yes, CaseSensitive=Yes, FollowedBy=TKG_SUBPROG_NAME)
    TKG_SUBPROG_NAME = \w[\w\d]+ (IsPattern=Yes, Restricted=Yes)
    TKG_EXTERN = EXTERN:\s (IsPattern=Yes, FollowedBy=TKG_PROG_FILE_NAME)
    TKG_PROG_FILE_NAME = [\^#&@']?[\w\d\./\:]+ (IsPattern=Yes, Restricted=Yes)
    TKG_PV_DECL = def:\s (IsPattern=Yes)
    TKG_PV_UNDECL = ~def:\s (IsPattern=Yes)
    TKG_VAR_RETAIN = retain:\s (IsPattern=Yes)
    TKG_VARSCOPE_IP_LOCAL = local:[\s\n] (IsPattern=Yes)
    TKG_VARSCOPE_IP_GLOBAL = ip_global:[\s\n] (IsPattern=Yes)
    TKG_VARSCOPE_NC_GLOBAL = nc_global:[\s\n] (IsPattern=Yes)
    TKG_VARSCOPE_PLC_GLOBAL = plc_global:[\s\n] (IsPattern=Yes)
    TKG_VARSYNCH_IP = ip_synch:\s (IsPattern=Yes)
    TKG_VARSYNCH_PATH = path_synch:\s (IsPattern=Yes)
    TKG_PAREVAL_DO = do:\s (FileXLInvalid=Yes, IsPattern=Yes)
    TKG_GOTOF = gotof:\s (FileXLInvalid=Yes, IsPattern=Yes, OptFollowedBy=TKG_GOTO_DEST)
    TKG_GOTOB = gotob:\s (FileXLInvalid=Yes, IsPattern=Yes, OptFollowedBy=TKG_GOTO_DEST)
    TKG_GOTO = goto:\s (FileXLInvalid=Yes, IsPattern=Yes, OptFollowedBy=TKG_GOTO_DEST)
    TKG_GOTO_DEST = \w[\w\d]* (IsPattern=Yes, Restricted=Yes)
    TKG_ARITH_BINARY_INT_DIVIDE = DIV:[\s(] (IsPattern=Yes)
    TKG_ARITH_BINARY_MODULO = MOD:[\s(] (IsPattern=Yes)
    TKG_FOR = FOR:\s (FileXLInvalid=Yes, IsPattern=Yes)
    TKG_ENDFOR = ENDFOR:[\s\n] (FileXLInvalid=Yes, IsPattern=Yes)
    TKG_FORTO = TO:\W (IsPattern=Yes)
    TKG_DO = repeat:[\s\n] (FileXLInvalid=Yes, IsPattern=Yes)
    TKG_ENDDO_UNTIL = until:[\s(] (FileXLInvalid=Yes, IsPattern=Yes)
    TKG_LOGICAL_UNARY_NOT = not:\W (IsPattern=Yes)
    TKG_SUPPRESS_SINGLE_STEP = NOHALT
    TKG_NC_BLOCK_PREFIX = N:[\s\d] (IsPattern=Yes)
    TKG_LOGICAL_HP_BINARY_AND = and:\W (IsPattern=Yes)
    TKG_LOGICAL_HP_BINARY_OR = or:\W (IsPattern=Yes)
    TKG_LOGICAL_HP_BINARY_XOR = xor:\W (IsPattern=Yes)
    TKG_BITWISE_BINARY_AND = b_and:\W (IsPattern=Yes)
    TKG_BITWISE_BINARY_OR = b_or:\W (IsPattern=Yes)
    TKG_BITWISE_BINARY_XOR = b_xor:\W (IsPattern=Yes)
    TKG_BITWISE_UNARY_COMPLEMENT = b_not:\W (IsPattern=Yes)
    TKG_PATHSYNCH_REC_IEC = do_path_synch:\W (FileXLInvalid=Yes, IsPattern=Yes)
    TKG_PATHSYNCH_END = end_path_synch:\W (FileXLInvalid=Yes, IsPattern=Yes)
    TKG_PATHSYNCH_IPEVAL = ip_eval:\W (FileXLInvalid=Yes, IsPattern=Yes)
    TKG_IF = if:\W (FileXLInvalid=Yes, IsPattern=Yes)
    TKG_THEN = then:\W (FileXLInvalid=Yes, IsPattern=Yes)
    TKG_BLOCK_ELSE = else:\W (FileXLInvalid=Yes, IsPattern=Yes)
    TKG_BLOCK_ENDIF = endif:\W (FileXLInvalid=Yes, IsPattern=Yes)
    TKG_SWITCH = case:\W (FileXLInvalid=Yes, IsPattern=Yes)
    TKG_SWITCH_OF = of:\W (FileXLInvalid=Yes, IsPattern=Yes)
    TKG_SWITCH_DEFAULT = default:\W (FileXLInvalid=Yes, IsPattern=Yes)
    TKG_WHILE = while:\W (FileXLInvalid=Yes, IsPattern=Yes)
    TKG_ENDWHILE = endwhile (FileXLInvalid=Yes)
    TKG_FOREVER = loop:\W (FileXLInvalid=Yes, IsPattern=Yes)
    TKG_ENDFOREVER = endloop:\W (FileXLInvalid=Yes, IsPattern=Yes)
    TKG_LABEL_DEF = \w:\:|\w[\w\d]+:\: (IsPattern=Yes, FollowedBy=TKG_LABEL_SUFFIX)
    TKG_LABEL_SUFFIX = : (Restricted=Yes)
    TKG_MACRO_TEXT = . (Restricted=Yes, IsPattern=Yes)
    TKG_MACRO_NAME = [$\w][$\w\d(]+ (Restricted=Yes, IsPattern=Yes)
    TKG_PRIM_TYPE (IsPattern=Yes)
    TKG_OPEN_BRACKET = (
    TKG_CLOSE_BRACKET = )
    TKG_OPEN_INDEXBRACKET = [
    TKG_CLOSE_INDEXBRACKET = ]
    TKG_COMMA = ,
    TKG_DOT = \.:\w (IsPattern=Yes, FollowedBy=TKG_STRUCT_MEMBER_REF)
    TKG_STRUCT_MEMBER_REF = \w|\w[\w\d]+ (IsPattern=Yes, Restricted=Yes)
    TKG_PARAM_PREFIX = R:[\[\d]|$[RP]:[\[\d]|M[WLF]:[\[\d]|EX[WLBF]:[\[\d] (IsPattern=Yes)
    TKG_SUBRANGE = ..
    TKG_NUMBER = \d+\.\d+|\d+\.:[^\.] (IsPattern=Yes)
    TKG_INTEGER = \d+ (IsPattern=Yes)
    TKG_FRACTION = \.\d+ (IsPattern=Yes)
    TKG_NUMBER_EXP = EX:[\s\d\+\-\.] (IsPattern=Yes)
    TKG_STRING_CONCAT = <<
    TKG_COMP_BINARY_GREATER_THAN_OR_EQ = >=
    TKG_COMP_BINARY_LESS_THAN_OR_EQ = <=
    TKG_COMP_BINARY_EQUAL_TO = ==
    TKG_COMP_BINARY_NOT_EQUAL_TO = <>
    TKG_COMP_BINARY_GREATER_THAN = >
    TKG_COMP_BINARY_LESS_THAN = <
    TKG_ASSIGN_INCR = =ic:( (IsPattern=Yes)
    TKG_ASSIGN_EQ = =
    TKG_ARITH_BINARY_PLUS = +
    TKG_ARITH_BINARY_MINUS = -
    TKG_ARITH_BINARY_MULTIPLY = *
    TKG_ARITH_BINARY_DIVIDE = /
    TKG_SUBCALL_REPEAT_PREFIX = P:[\s\d] (IsPattern=Yes, FollowedBy=TKG_INTEGER)
    TKG_PV_DECL_REF = \w[\w\d\.\:\*]* (IsPattern=Yes, Restricted=Yes)
    TKG_G_CODE_PREFIX = G:[\s\d] (IsPattern=Yes)
    TKG_M_CODE_PREFIX = M:[\s\d(] (IsPattern=Yes)
    TKG_FUB_DECL = fub\s (IsPattern=Yes)
    TKG_FUB_ERR_LEV_1 = error_level_1:\s (IsPattern=Yes)
    TKG_FUB_ERR_LEV_2 = error_level_2:\s (IsPattern=Yes)
    TKG_FUB_ERR_LEV_3 = error_level_3:\s (IsPattern=Yes)
    TKG_FUB_ERR_LEV_4 = error_level_4:\s (IsPattern=Yes)
    TKG_FUB_BLOCKING = blocking:[\s\n] (IsPattern=Yes)
    TKG_FUB_NON_BLOCKING = non_blocking:\s (IsPattern=Yes)
    TKG_IEC_TYPED_VALUE = #[\w\d]+:[^\w\d\:] (IsPattern=Yes)
    TKG_REFERENCE = ref:[\s\n]|reference:[\s\n] (IsPattern=Yes, FollowedBy=TKG_IEC_TO)
    TKG_IEC_TO = to:[\s\n] (IsPattern=Yes, Restricted=Yes)
    TKG_ACCESS = ACCESS:[\s\n] (IsPattern=Yes)
    TKG_BINARY_LITERAL_START = 'B:[01_] (FollowedBy=TKG_BINARY_LITERAL_BODY, IsPattern=Yes)
    TKG_BINARY_LITERAL_BODY = [01_]+' (Restricted=Yes, IsPattern=Yes)
    TKG_HEX_LITERAL_START = 'H:[\dA-F_] (FollowedBy=TKG_HEX_LITERAL_BODY, IsPattern=Yes)
    TKG_HEX_LITERAL_BODY = [\dA-F_]+' (Restricted=Yes, IsPattern=Yes)
    TKG_WORD = \w|\w[\w\d\./]+|\./\w|\./\w[\w\d\./]+|[\^#][\w\d]+\:[\w\d\./]+ (IsPattern=Yes)
  StringChars (AsciiStringStart=", AsciiStringEnd=", UTF16StringStart=W", UTF16StringEnd=")
    EscapeSeq (Search=$N, ReplaceValue=10)
    EscapeSeq (Search=$L, ReplaceValue=10)
    EscapeSeq (Search=$P, ReplaceValue=12)
    EscapeSeq (Search=$R, ReplaceValue=13)
    EscapeSeq (Search=$T, ReplaceValue=9)
    EscapeSeq (Search=$Q, ReplaceStr=")
    EscapeSeq (Search=$', ReplaceStr=')
    EscapeSeq (Search=$", ReplaceStr=")
    EscapeSeq (Search=$[\dA-Fa-f]+, IsPattern=Yes, ReplaceEncodingBase=16)
    EscapeSeq (Search=$$, ReplaceStr=$)
    EscapeSeq (Search=$, ReplaceStr=)
```

### Data object Logical/GmcIpConfig/gmcipcsm (Cnc, version 5.02.1)

#### gmcipcsm.cnc
```
Root (LangModule=ailgcode, Version=1.0)
  Constants:
    NumAxes = 15 (Type=INT)
  Preprocess:
    PP_RULE_STOPRE (Search=STOPRE, Replace=G172)
    PP_RULE_CIP (Search=CIP:\W, Replace=G102, IsPattern=Yes)
  Types:
    RotationAngleSpecifier (type=ENUM, EnumType=REGEXP, Value6=H)
    RadiusSpecifier (type=ENUM, EnumType=REGEXP, Value1=R\s*=, Value2=CR\s*=)
    InterpolParam (type=ENUM, EnumType=REGEXP, Value0=I, Value1=J, Value2=K, Value100=G161\s*I, Value101=G161\s*J, Value102=G161\s*K, Value200=G162\s*I, Value201=G162\s*J, Value202=G162\s*K, Value0300=I\s*=\s*AC, Value0301=J\s*=\s*AC, Value0302=K\s*=\s*AC, Value0400=I\s*=\s*IC, Value0401=J\s*=\s*IC, Value0402=K\s*=\s*IC)
    CirclePointParam (type=ENUM, EnumType=REGEXP, Value0=I1\s*=, Value1=J1\s*=, Value2=K1\s*=, Value100=G161\s*I1\s*=, Value101=G161\s*J1\s*=, Value102=G161\s*K1\s*=, Value200=G162\s*I1\s*=, Value201=G162\s*J1\s*=, Value202=G162\s*K1\s*=, Value0300=I1\s*=\s*AC, Value0301=J1\s*=\s*AC, Value0302=K1\s*=\s*AC, Value0400=I1\s*=\s*IC, Value0401=J1\s*=\s*IC, Value0402=K1\s*=\s*IC)
    RPYAngleName (type=ENUM, EnumType=REGEXP, Value1=ROLL, Value0=PITCH, Value2=YAW)
    EulerAngleName (type=ENUM, EnumType=REGEXP, Value3=PHI, Value4=THETA, Value5=PSI)
    RotaryVectorName (type=ENUM, EnumType=REGEXP, Value0=P\s*=, Value1=Q\s*=, Value2=R\s*=)
    DwellTime (type=FLOAT)
    RParamIndex (type=INT, MinValue=0, MaxValue=999)
    EXParamIndex (type=INT, MinValue=0, MaxValue=99)
    MParamIndex (type=INT, MinValue=0, MaxValue=99)
    Byte (type=INT, MinValue=0, MaxValue=255)
    Word (type=INT, MinValue=-32768, MaxValue=32767)
    Long (type=INT)
  PVMacros:
    SAVE (ArrayDims=0, Group=500)
      CALL = Info(:id:52101, msg:"Save Modal GCode State NOT SUPPORTED YET":);
  SysVars
  Parameters:
    R (IndexType=RParamIndex, ValueType=FLOAT)
      ARG (ref=EXPR, DataType=RParamIndex)
    QUOTED (QuotedName=$R, Synchronous=Yes, IndexType=RParamIndex, ValueType=FLOAT)
      ARG (ref=EXPR, DataType=RParamIndex)
    QUOTED (QuotedName=$P, Synchronous=Yes, IndexType=RParamIndex, ValueType=FLOAT)
      ARG (ref=EXPR, DataType=RParamIndex)
    EXB (IndexType=EXParamIndex, ValueType=Byte)
      ARG (ref=EXPR, DataType=EXParamIndex)
    EXW (IndexType=EXParamIndex, ValueType=Word)
      ARG (ref=EXPR, DataType=EXParamIndex)
    EXL (IndexType=EXParamIndex, ValueType=Long)
      ARG (ref=EXPR, DataType=EXParamIndex)
    EXF (IndexType=EXFParamIndex, ValueType=FLOAT)
      ARG (ref=EXPR, DataType=EXFParamIndex)
    MW (Synchronous=Yes, IndexType=MParamIndex, ValueType=Word)
      ARG (ref=EXPR, DataType=MParamIndex)
    ML (Synchronous=Yes, IndexType=MParamIndex, ValueType=Long)
      ARG (ref=EXPR, DataType=MParamIndex)
    MF (Synchronous=Yes, IndexType=MParamIndex, ValueType=FLOAT)
      ARG (ref=EXPR, DataType=MParamIndex)
  MCodes:
    M17 = 17 (Group=41, Alias=RET:[^\d\w\(], Eval=Early, Inline=Yes, AliasIsPattern=Yes)
      ARG (ref=VALUE, DataType=FLOAT, RequireLiteral=Yes)
    M17_1 = 17.1 (Group=41, Alias=CONDRET, Eval=Early, Inline=Yes)
      ARG (ref=VALUE, DataType=FLOAT, RequireLiteral=Yes)
```

### Data object Logical/GmcIpConfig/gmcipcfg (Cnc, version 5.02.1)

#### gmcipcfg.cnc
```
CONFIG:
  LANG_INCLUDE gmcipmxd (LangName=IEC-ST, DataObject=Yes, IfNotExist=Error, Scope=NC_GLOBAL, RequireFnIgnore=MXConvertOrient)
  XML_INCLUDE gmcipvar (IfNotExist=Warn)
  XML_INCLUDE gmcipfun (IfNotExist=Warn)
  XML_INCLUDE gmcipfub (IfNotExist=Warn)
  MPQUEUE (NumPackets=200, LookaheadMinBlocks=5, LookaheadMaxBlocks=20, LookaheadMode=any, MaxPathJobs=256, CheckForNaNs=1)
  MONITOR (MaxPathStackEvents=1024)
  MPLOG (MaxBuffers=10, MinBuffers=4, EarlyCircleBufferLookahead=2, DefaultBufferSize=131072, TaskCycleDelay=1, FileDevice=mplog*, MaxLogFiles=20, MaxLogFileSize=1048576, CopyLineTextMaxChars=80)
  AXES (StandardCNCAxes=Yes)
  FUBOutputs:
    FUBOutput PLCOpen:
      ERROR (condition=$Error == 1)
      BUSY (condition=$Busy == 1)
    FUBOutput BuR:
      ERROR (condition=$status != 65535 && $status != 0)
      BUSY (condition=$status == 65535)
  FUNCTIONS:
    FUNC LEN (DeclareName=__LEN, AlwaysDeclare=Yes, RetType=INT)
      ARG IN (Type=STRING)
    FUNC LEFT (DeclareName=__LEFT, AlwaysDeclare=Yes, RetType=STRING, RetRef=Yes)
      ARG IN (Type=STRING)
      ARG L (Type=INT)
    FUNC RIGHT (DeclareName=__RIGHT, AlwaysDeclare=Yes, RetType=STRING, RetRef=Yes)
      ARG IN (Type=STRING)
      ARG L (Type=INT)
    FUNC MID (DeclareName=__MID, AlwaysDeclare=Yes, RetType=STRING, RetRef=Yes)
      ARG IN (Type=STRING)
      ARG L (Type=INT)
      ARG P (Type=INT)
    FUNC CONCAT (DeclareName=__CONCAT, AlwaysDeclare=Yes, RetType=STRING, RetRef=Yes)
      ARG IN1 (Type=STRING)
      ARG IN2 (Type=STRING)
    FUNC INSERT (DeclareName=__INSERT, AlwaysDeclare=Yes, RetType=STRING, RetRef=Yes)
      ARG IN1 (Type=STRING)
      ARG IN2 (Type=STRING)
      ARG P (Type=INT)
    FUNC DELETE (DeclareName=__DELETE, AlwaysDeclare=Yes, RetType=STRING, RetRef=Yes)
      ARG IN (Type=STRING)
      ARG L (Type=INT)
      ARG P (Type=INT)
    FUNC REPLACE (DeclareName=__REPLACE, AlwaysDeclare=Yes, RetType=STRING, RetRef=Yes)
      ARG IN1 (Type=STRING)
      ARG IN2 (Type=STRING)
      ARG L (Type=INT)
      ARG P (Type=INT)
    FUNC FIND (DeclareName=__FIND, AlwaysDeclare=Yes, RetType=INT)
      ARG IN1 (Type=STRING)
      ARG IN2 (Type=STRING)
  XML_INCLUDE gmcipuc (IfNotExist=Warn)
```

### Data object Logical/GmcIpConfig/gmcipiec (Cnc, version 5.02.1)

#### gmcipiec.cnc
```
Root (LangModule=ailgcode, Version=1.0)
  AxesSpec
  PrimTypes (PatternSuffix=:[^\d\w$#])
    BOOL (BRType=BOOL)
    STRING (BRType=STRING)
    WSTRING (BRType=WSTRING)
    TIME (BRType=TIME)
    SINT (BRType=SINT)
    INT (BRType=INT)
    DINT (BRType=DINT)
    USINT (BRType=USINT)
    UINT (BRType=UINT)
    UDINT (BRType=UDINT)
    REAL (BRType=REAL)
    LREAL (BRType=LREAL)
    DATE (BRType=DATE)
    DATE_AND_TIME (BRType=DATE_AND_TIME)
    DT (BRType=DT)
    TIME_OF_DAY (BRType=TIME_OF_DAY)
    TOD (BRType=TIME_OF_DAY)
    BYTE (BRType=BYTE)
    WORD (BRType=WORD)
    DWORD (BRType=DWORD)
  BuiltInProcs:
    SetCyclicId = #job->group_id = $[1]; (MinArgs=1, MaxArgs=1, Eval=Early)
    WaitForCyclic = if ( Defined(:$[1]:) ) 
        WaitForCyclicGroups(:${*}:);  
      else
        WaitForCyclicJob(:#last_job_id:);
      endif (MinArgs=0, MaxArgs=*)
    REPORT (MinArgs=2, MaxArgs=2)
      Arg (ref=id, DataType=INT)
      Arg (ref=msg, DataType=STRING)
    WARN (MinArgs=2, MaxArgs=2)
      Arg (ref=id, DataType=INT)
      Arg (ref=msg, DataType=STRING)
    HALT (MinArgs=2, MaxArgs=2)
      Arg (ref=id, DataType=INT)
      Arg (ref=msg, DataType=STRING)
    ERROR (MinArgs=2, MaxArgs=2)
      Arg (ref=id, DataType=INT)
      Arg (ref=msg, DataType=STRING)
    LOADBG (MinArgs=1, MaxArgs=1)
      Arg (ref=filename, DataType=STRING)
    LOAD (MinArgs=1, MaxArgs=1)
      Arg (ref=filename, DataType=STRING)
    UNLOAD (MinArgs=1, MaxArgs=1)
      Arg (ref=filename, DataType=STRING)
    EXEC (MinArgs=1, MaxArgs=5)
      Arg (ref=filename, DataType=STRING)
      Arg (ref=arguments, DataType=ANY_DATA)
      Arg (ref=langId, DataType=INT)
      Arg (ref=block, DataType=INT, MinCount=0, MaxCount=1, DenyArgs=5, WriteOpts=:)
      Arg (ref=line, DataType=INT, MinCount=0, MaxCount=1, DenyArgs=4, WriteOpts=:)
    EXEC_RPC (MinArgs=2, MaxArgs=4)
      Arg (ref=filename, DataType=STRING)
      Arg (ref=arguments, DataType=ANY_DATA)
      Arg (ref=langId, DataType=INT)
      Arg (ref=rpc, DataType=ANY_DATA, MinCount=1, MaxCount=1)
    EVAL (MinArgs=1, MaxArgs=2)
      Arg (ref=expression, DataType=STRING)
      Arg (ref=langId, DataType=INT)
    PUSH_PACKET = PushPacket(::);
    PUSH_PACKET_CMD (MinArgs=1, MaxArgs=2)
      Arg (ref=cmd, DataType=INT)
      Arg (ref=data, DataType=ANY_DATA)
    DISPATCH_AND_WAIT (MinArgs=1, MaxArgs=1)
      Arg (ref=cmd, DataType=INT)
    START_PACKET_LIST = #inhibit_mp_list_dispatch = 1;
    END_PACKET_LIST = #inhibit_mp_list_dispatch = 0;
    LOG_INFO (MinArgs=1, MaxArgs=1)
      Arg (ref=msg, DataType=STRING)
    SET_BLOCK_NUMBER = SetCurBlockNr(:$[1]:); (MinArgs=1, MaxArgs=1)
    SBLOF_PATH = #next_motion.Command = MPCMD_SBL_PATH_INHIBIT;
      PushPacket(::);
    SBLON_PATH = #next_motion.Command = MPCMD_SBL_PATH_RELEASE;
      PushPacket(::);
  BuiltInFns:
    ABS = Abs(:$[1]:) (ReturnType=ANY_NUM, ArgType1=ANY_NUM, Inline=Yes)
    SIN = RSin(:$[1]:) (ReturnType=ANY_REAL, ArgType1=ANY_REAL, Inline=Yes)
    COS = RCos(:$[1]:) (ReturnType=ANY_REAL, ArgType1=ANY_REAL, Inline=Yes)
    TAN = RTan(:$[1]:) (ReturnType=ANY_REAL, ArgType1=ANY_REAL, Inline=Yes)
    ASIN = RASin(:$[1]:) (ReturnType=ANY_REAL, ArgType1=ANY_REAL, Inline=Yes)
    ACOS = RACos(:$[1]:) (ReturnType=ANY_REAL, ArgType1=ANY_REAL, Inline=Yes)
    ATAN = RATan(:$[1]:) (ReturnType=ANY_REAL, ArgType1=ANY_REAL, Inline=Yes)
    SQRT = Sqrt(:$[1]:) (ReturnType=ANY_REAL, ArgType1=ANY_REAL, Inline=Yes)
    LN = Ln(:$[1]:) (ReturnType=ANY_REAL, ArgType1=ANY_REAL, Inline=Yes)
    EXP = Exp(:$[1]:) (ReturnType=ANY_REAL, ArgType1=ANY_REAL, Inline=Yes)
    LOG = Log(:$[1]:) (ReturnType=ANY_REAL, ArgType1=ANY_REAL, Inline=Yes)
    EXPT = Pow(:$[1],$[2]:) (ReturnType=ANY_REAL, ArgType1=ANY_REAL, ArgType2=ANY_NUM, Inline=Yes)
    TRUNC = ToInt(:Fix(:$[1]:):) (ReturnType=IEC_INT, ArgType1=ANY_REAL, Inline=Yes)
    ADR = Adr(:\$[1]:) (ReturnType=IEC_UDINT, ArgType1=ANY_DATA, Inline=Yes)
    REF = \$[1] (ReturnType=ANY_DATA, ArgType1=ANY_DATA, Inline=Yes)
    SIZEOF = Sizeof(:\$[1]:) (ReturnType=IEC_UINT, NumArgs=1, Inline=Yes)
    LIMIT (ReturnType=ANY_NUM, Inline=No)
      Arg (ref=MIN, DataType=ANY_NUM)
      Arg (ref=IN, DataType=ANY_NUM)
      Arg (ref=MAX, DataType=ANY_NUM)
    MIN (ReturnType=ANY_NUM, Inline=No)
      Arg (ref=IN1, DataType=ANY_NUM)
      Arg (ref=IN2, DataType=ANY_NUM)
    MAX (ReturnType=ANY_NUM, Inline=No)
      Arg (ref=IN1, DataType=ANY_NUM)
      Arg (ref=IN2, DataType=ANY_NUM)
    ROL = BitRotL(:$[1],$[2]:) (ReturnType=ANY_NUM, ArgType1=ANY_NUM, ArgType2=IEC_SINT)
    ROR = BitRotR(:$[1],$[2]:) (ReturnType=ANY_NUM, ArgType1=ANY_NUM, ArgType2=IEC_SINT)
    SHR = BitShR(:$[1],$[2]:) (ReturnType=ANY_NUM, ArgType1=ANY_NUM, ArgType2=IEC_SINT)
    SHL = BitShL(:$[1],$[2]:) (ReturnType=ANY_NUM, ArgType1=ANY_NUM, ArgType2=IEC_SINT)
    BIT_TST = AsBitTst(:$[1],$[2]:) (ReturnType=ANY_NUM, ArgType1=ANY_NUM, ArgType2=IEC_SINT)
    BIT_SET = AsBitSet(:$[1],$[2]:) (ReturnType=ANY_NUM, ArgType1=ANY_NUM, ArgType2=IEC_SINT)
    BIT_CLR = AsBitClr(:$[1],$[2]:) (ReturnType=ANY_NUM, ArgType1=ANY_NUM, ArgType2=IEC_SINT)
    TO_BOOL = ToBool(:$[1]:) (ReturnType=IEC_BOOL, ArgType1=ANY_DATA, Inline=Yes)
    TO_USINT = ToUInt(:$[1],1:) (ReturnType=IEC_USINT, ArgType1=ANY_DATA, Inline=Yes)
    TO_BYTE = ToUInt(:$[1],1:) (ReturnType=IEC_BYTE, ArgType1=ANY_DATA, Inline=Yes)
    TO_SINT = ToInt(:$[1],1:) (ReturnType=IEC_SINT, ArgType1=ANY_DATA, Inline=Yes)
    TO_UINT = ToUInt(:$[1],2:) (ReturnType=IEC_UINT, ArgType1=ANY_DATA, Inline=Yes)
    TO_WORD = ToUInt(:$[1],2:) (ReturnType=IEC_WORD, ArgType1=ANY_DATA, Inline=Yes)
    TO_INT = ToInt(:$[1],2:) (ReturnType=IEC_INT, ArgType1=ANY_DATA, Inline=Yes)
    TO_UDINT = ToUInt(:$[1]:) (ReturnType=IEC_UDINT, ArgType1=ANY_DATA, Inline=Yes)
    TO_DWORD = ToUInt(:$[1]:) (ReturnType=IEC_DWORD, ArgType1=ANY_DATA, Inline=Yes)
    TO_DINT = ToInt(:$[1]:) (ReturnType=IEC_DINT, ArgType1=ANY_DATA, Inline=Yes)
    TO_TIME = ToTime(:$[1]:) (ReturnType=IEC_TIME, ArgType1=ANY_DATA, Inline=Yes)
    TO_DT = ToDT(:$[1]:) (ReturnType=IEC_DT, ArgType1=ANY_DATA, Inline=Yes)
    TO_DATE_AND_TIME = ToDT(:$[1]:) (ReturnType=IEC_DT, ArgType1=ANY_DATA, Inline=Yes)
    TO_TOD = ToTOD(:$[1]:) (ReturnType=IEC_TOD, ArgType1=ANY_DATA, Inline=Yes)
    TO_TIME_OF_DAY = ToTOD(:$[1]:) (ReturnType=IEC_TOD, ArgType1=ANY_DATA, Inline=Yes)
    TO_DATE = ToDate(:$[1]:) (ReturnType=IEC_DATE, ArgType1=ANY_DATA, Inline=Yes)
    TO_REAL = ToFloat(:$[1]:) (ReturnType=IEC_REAL, ArgType1=ANY_DATA, Inline=Yes)
    TO_LREAL = ToLReal(:$[1]:) (ReturnType=IEC_LREAL, ArgType1=ANY_DATA, Inline=Yes)
    TO_STRING = ToString(:$[1]:) (ReturnType=IEC_STRING, ArgType1=ANY_DATA, Inline=Yes)
    TO_WSTRING = ToWString(:$[1]:) (ReturnType=IEC_WSTRING, ArgType1=ANY_DATA, Inline=Yes)
    USINT_TO_BOOL = ToBool(:$[1]:) (ReturnType=IEC_BOOL, ArgType1=IEC_USINT, Inline=Yes)
    SINT_TO_BOOL = ToBool(:$[1]:) (ReturnType=IEC_BOOL, ArgType1=IEC_SINT, Inline=Yes)
    UINT_TO_BOOL = ToBool(:$[1]:) (ReturnType=IEC_BOOL, ArgType1=IEC_UINT, Inline=Yes)
    INT_TO_BOOL = ToBool(:$[1]:) (ReturnType=IEC_BOOL, ArgType1=IEC_INT, Inline=Yes)
    UDINT_TO_BOOL = ToBool(:$[1]:) (ReturnType=IEC_BOOL, ArgType1=IEC_UDINT, Inline=Yes)
    DINT_TO_BOOL = ToBool(:$[1]:) (ReturnType=IEC_BOOL, ArgType1=IEC_DINT, Inline=Yes)
    REAL_TO_BOOL = ToBool(:$[1]:) (ReturnType=IEC_BOOL, ArgType1=IEC_REAL, Inline=Yes)
    LREAL_TO_BOOL = ToBool(:$[1]:) (ReturnType=IEC_BOOL, ArgType1=IEC_LREAL, Inline=Yes)
    TIME_TO_BOOL = ToBool(:$[1]:) (ReturnType=IEC_BOOL, ArgType1=IEC_TIME, Inline=Yes)
    DT_TO_BOOL = ToBool(:$[1]:) (ReturnType=IEC_BOOL, ArgType1=IEC_DT, Inline=Yes)
    TOD_TO_BOOL = ToBool(:$[1]:) (ReturnType=IEC_BOOL, ArgType1=IEC_TOD, Inline=Yes)
    BYTE_TO_BOOL = ToBool(:$[1]:) (ReturnType=IEC_BOOL, ArgType1=IEC_BYTE, Inline=Yes)
    WORD_TO_BOOL = ToBool(:$[1]:) (ReturnType=IEC_BOOL, ArgType1=IEC_WORD, Inline=Yes)
    DWORD_TO_BOOL = ToBool(:$[1]:) (ReturnType=IEC_BOOL, ArgType1=IEC_DWORD, Inline=Yes)
    BOOL_TO_USINT = ToUInt(:$[1],1:) (ReturnType=IEC_USINT, ArgType1=IEC_BOOL, Inline=Yes)
    SINT_TO_USINT = ToUInt(:$[1],1:) (ReturnType=IEC_USINT, ArgType1=IEC_SINT, Inline=Yes)
    UINT_TO_USINT = ToUInt(:$[1],1:) (ReturnType=IEC_USINT, ArgType1=IEC_UINT, Inline=Yes)
    INT_TO_USINT = ToUInt(:$[1],1:) (ReturnType=IEC_USINT, ArgType1=IEC_INT, Inline=Yes)
    UDINT_TO_USINT = ToUInt(:$[1],1:) (ReturnType=IEC_USINT, ArgType1=IEC_UDINT, Inline=Yes)
    DINT_TO_USINT = ToUInt(:$[1],1:) (ReturnType=IEC_USINT, ArgType1=IEC_DINT, Inline=Yes)
    REAL_TO_USINT = ToUInt(:$[1],1:) (ReturnType=IEC_USINT, ArgType1=IEC_REAL, Inline=Yes)
    LREAL_TO_USINT = ToUInt(:$[1],1:) (ReturnType=IEC_USINT, ArgType1=IEC_LREAL, Inline=Yes)
    BOOL_TO_SINT = ToInt(:$[1],1:) (ReturnType=IEC_SINT, ArgType1=IEC_BOOL, Inline=Yes)
    USINT_TO_SINT = ToInt(:$[1],1:) (ReturnType=IEC_SINT, ArgType1=IEC_USINT, Inline=Yes)
    UINT_TO_SINT = ToInt(:$[1],1:) (ReturnType=IEC_SINT, ArgType1=IEC_UINT, Inline=Yes)
    INT_TO_SINT = ToInt(:$[1],1:) (ReturnType=IEC_SINT, ArgType1=IEC_INT, Inline=Yes)
    UDINT_TO_SINT = ToInt(:$[1],1:) (ReturnType=IEC_SINT, ArgType1=IEC_UDINT, Inline=Yes)
    DINT_TO_SINT = ToInt(:$[1],1:) (ReturnType=IEC_SINT, ArgType1=IEC_DINT, Inline=Yes)
    REAL_TO_SINT = ToInt(:$[1],1:) (ReturnType=IEC_SINT, ArgType1=IEC_REAL, Inline=Yes)
    LREAL_TO_SINT = ToInt(:$[1],1:) (ReturnType=IEC_SINT, ArgType1=IEC_LREAL, Inline=Yes)
    BOOL_TO_UINT = ToUInt(:$[1],2:) (ReturnType=IEC_UINT, ArgType1=IEC_BOOL, Inline=Yes)
    SINT_TO_UINT = ToUInt(:$[1],2:) (ReturnType=IEC_UINT, ArgType1=IEC_SINT, Inline=Yes)
    USINT_TO_UINT = ToUInt(:$[1],2:) (ReturnType=IEC_UINT, ArgType1=IEC_USINT, Inline=Yes)
    INT_TO_UINT = ToUInt(:$[1],2:) (ReturnType=IEC_UINT, ArgType1=IEC_INT, Inline=Yes)
    UDINT_TO_UINT = ToUInt(:$[1],2:) (ReturnType=IEC_UINT, ArgType1=IEC_UDINT, Inline=Yes)
    DINT_TO_UINT = ToUInt(:$[1],2:) (ReturnType=IEC_UINT, ArgType1=IEC_DINT, Inline=Yes)
    REAL_TO_UINT = ToUInt(:$[1],2:) (ReturnType=IEC_UINT, ArgType1=IEC_REAL, Inline=Yes)
    LREAL_TO_UINT = ToUInt(:$[1],2:) (ReturnType=IEC_UINT, ArgType1=IEC_LREAL, Inline=Yes)
    BOOL_TO_INT = ToInt(:$[1],2:) (ReturnType=IEC_INT, ArgType1=IEC_BOOL, Inline=Yes)
    SINT_TO_INT = ToInt(:$[1],2:) (ReturnType=IEC_INT, ArgType1=IEC_SINT, Inline=Yes)
    USINT_TO_INT = ToInt(:$[1],2:) (ReturnType=IEC_INT, ArgType1=IEC_USINT, Inline=Yes)
    UINT_TO_INT = ToInt(:$[1],2:) (ReturnType=IEC_INT, ArgType1=IEC_UINT, Inline=Yes)
    UDINT_TO_INT = ToInt(:$[1],2:) (ReturnType=IEC_INT, ArgType1=IEC_UDINT, Inline=Yes)
    DINT_TO_INT = ToInt(:$[1],2:) (ReturnType=IEC_INT, ArgType1=IEC_DINT, Inline=Yes)
    REAL_TO_INT = ToInt(:$[1],2:) (ReturnType=IEC_INT, ArgType1=IEC_REAL, Inline=Yes)
    LREAL_TO_INT = ToInt(:$[1],2:) (ReturnType=IEC_INT, ArgType1=IEC_LREAL, Inline=Yes)
    BOOL_TO_UDINT = ToUInt(:$[1]:) (ReturnType=IEC_UDINT, ArgType1=IEC_BOOL, Inline=Yes)
    USINT_TO_UDINT = ToUInt(:$[1]:) (ReturnType=IEC_UDINT, ArgType1=IEC_USINT, Inline=Yes)
    SINT_TO_UDINT = ToUInt(:$[1]:) (ReturnType=IEC_UDINT, ArgType1=IEC_SINT, Inline=Yes)
    UINT_TO_UDINT = ToUInt(:$[1]:) (ReturnType=IEC_UDINT, ArgType1=IEC_UINT, Inline=Yes)
    INT_TO_UDINT = ToUInt(:$[1]:) (ReturnType=IEC_UDINT, ArgType1=IEC_INT, Inline=Yes)
    DINT_TO_UDINT = ToUInt(:$[1]:) (ReturnType=IEC_UDINT, ArgType1=IEC_DINT, Inline=Yes)
    REAL_TO_UDINT = ToUInt(:$[1]:) (ReturnType=IEC_UDINT, ArgType1=IEC_REAL, Inline=Yes)
    LREAL_TO_UDINT = ToUInt(:$[1]:) (ReturnType=IEC_UDINT, ArgType1=IEC_LREAL, Inline=Yes)
    TIME_TO_UDINT = ToUInt(:$[1]:) (ReturnType=IEC_UDINT, ArgType1=IEC_TIME, Inline=Yes)
    DT_TO_UDINT = ToUInt(:$[1]:) (ReturnType=IEC_UDINT, ArgType1=IEC_DT, Inline=Yes)
    BOOL_TO_DINT = ToInt(:$[1]:) (ReturnType=IEC_DINT, ArgType1=IEC_BOOL, Inline=Yes)
    USINT_TO_DINT = ToInt(:$[1]:) (ReturnType=IEC_DINT, ArgType1=IEC_USINT, Inline=Yes)
    SINT_TO_DINT = ToInt(:$[1]:) (ReturnType=IEC_DINT, ArgType1=IEC_SINT, Inline=Yes)
    UINT_TO_DINT = ToInt(:$[1]:) (ReturnType=IEC_DINT, ArgType1=IEC_UINT, Inline=Yes)
    INT_TO_DINT = ToInt(:$[1]:) (ReturnType=IEC_DINT, ArgType1=IEC_INT, Inline=Yes)
    UDINT_TO_DINT = ToInt(:$[1]:) (ReturnType=IEC_DINT, ArgType1=IEC_UDINT, Inline=Yes)
    REAL_TO_DINT = ToInt(:$[1]:) (ReturnType=IEC_DINT, ArgType1=IEC_REAL, Inline=Yes)
    LREAL_TO_DINT = ToInt(:$[1]:) (ReturnType=IEC_DINT, ArgType1=IEC_LREAL, Inline=Yes)
    TIME_TO_DINT = ToInt(:$[1]:) (ReturnType=IEC_DINT, ArgType1=IEC_TIME, Inline=Yes)
    DT_TO_DINT = ToInt(:$[1]:) (ReturnType=IEC_DINT, ArgType1=IEC_DT, Inline=Yes)
    BOOL_TO_TIME = ToTime(:$[1]:) (ReturnType=IEC_TIME, ArgType1=IEC_BOOL, Inline=Yes)
    DINT_TO_TIME = ToTime(:$[1]:) (ReturnType=IEC_TIME, ArgType1=IEC_DINT, Inline=Yes)
    UDINT_TO_TIME = ToTime(:$[1]:) (ReturnType=IEC_TIME, ArgType1=IEC_UDINT, Inline=Yes)
    BOOL_TO_DT = ToDT(:$[1]:) (ReturnType=IEC_DT, ArgType1=IEC_BOOL, Inline=Yes)
    DINT_TO_DT = ToDT(:$[1]:) (ReturnType=IEC_DT, ArgType1=IEC_DINT, Inline=Yes)
    UDINT_TO_DT = ToDT(:$[1]:) (ReturnType=IEC_DT, ArgType1=IEC_UDINT, Inline=Yes)
    BOOL_TO_REAL = ToFloat(:$[1]:) (ReturnType=IEC_REAL, ArgType1=IEC_BOOL, Inline=Yes)
    USINT_TO_REAL = ToFloat(:$[1]:) (ReturnType=IEC_REAL, ArgType1=IEC_USINT, Inline=Yes)
    SINT_TO_REAL = ToFloat(:$[1]:) (ReturnType=IEC_REAL, ArgType1=IEC_SINT, Inline=Yes)
    UINT_TO_REAL = ToFloat(:$[1]:) (ReturnType=IEC_REAL, ArgType1=IEC_UINT, Inline=Yes)
    INT_TO_REAL = ToFloat(:$[1]:) (ReturnType=IEC_REAL, ArgType1=IEC_INT, Inline=Yes)
    UDINT_TO_REAL = ToFloat(:$[1]:) (ReturnType=IEC_REAL, ArgType1=IEC_UDINT, Inline=Yes)
    DINT_TO_REAL = ToFloat(:$[1]:) (ReturnType=IEC_REAL, ArgType1=IEC_DINT, Inline=Yes)
    LREAL_TO_REAL = ToFloat(:$[1]:) (ReturnType=IEC_REAL, ArgType1=IEC_LREAL, Inline=Yes)
    TIME_TO_REAL = ToFloat(:$[1]:) (ReturnType=IEC_REAL, ArgType1=IEC_TIME, Inline=Yes)
    BOOL_TO_LREAL = ToLReal(:$[1]:) (ReturnType=IEC_LREAL, ArgType1=IEC_BOOL, Inline=Yes)
    USINT_TO_LREAL = ToLReal(:$[1]:) (ReturnType=IEC_LREAL, ArgType1=IEC_USINT, Inline=Yes)
    SINT_TO_LREAL = ToLReal(:$[1]:) (ReturnType=IEC_LREAL, ArgType1=IEC_SINT, Inline=Yes)
    UINT_TO_LREAL = ToLReal(:$[1]:) (ReturnType=IEC_LREAL, ArgType1=IEC_UINT, Inline=Yes)
    INT_TO_LREAL = ToLReal(:$[1]:) (ReturnType=IEC_LREAL, ArgType1=IEC_INT, Inline=Yes)
    UDINT_TO_LREAL = ToLReal(:$[1]:) (ReturnType=IEC_LREAL, ArgType1=IEC_UDINT, Inline=Yes)
    DINT_TO_LREAL = ToLReal(:$[1]:) (ReturnType=IEC_LREAL, ArgType1=IEC_DINT, Inline=Yes)
    REAL_TO_LREAL = ToLReal(:$[1]:) (ReturnType=IEC_LREAL, ArgType1=IEC_REAL, Inline=Yes)
    TIME_TO_LREAL = ToLReal(:$[1]:) (ReturnType=IEC_LREAL, ArgType1=IEC_TIME, Inline=Yes)
    BOOL_TO_STRING = ToString(:ToBool(:$[1]:):) (ReturnType=IEC_STRING, ArgType1=IEC_BOOL, Inline=Yes)
    USINT_TO_STRING = ToString(:ToUInt(:$[1],1:):) (ReturnType=IEC_STRING, ArgType1=IEC_USINT, Inline=Yes)
    SINT_TO_STRING = ToString(:ToInt(:$[1],1:):) (ReturnType=IEC_STRING, ArgType1=IEC_SINT, Inline=Yes)
    UINT_TO_STRING = ToString(:ToUInt(:$[1],2:):) (ReturnType=IEC_STRING, ArgType1=IEC_UINT, Inline=Yes)
    INT_TO_STRING = ToString(:ToInt(:$[1],2:):) (ReturnType=IEC_STRING, ArgType1=IEC_INT, Inline=Yes)
    UDINT_TO_STRING = ToString(:ToUInt(:$[1]:):) (ReturnType=IEC_STRING, ArgType1=IEC_UDINT, Inline=Yes)
    DINT_TO_STRING = ToString(:ToInt(:$[1]:):) (ReturnType=IEC_STRING, ArgType1=IEC_DINT, Inline=Yes)
    REAL_TO_STRING = ToString(:ToFloat(:$[1]:):) (ReturnType=IEC_STRING, ArgType1=IEC_REAL, Inline=Yes)
    LREAL_TO_STRING = ToString(:ToLReal(:$[1]:):) (ReturnType=IEC_STRING, ArgType1=IEC_LREAL, Inline=Yes)
    STRING_TO_BOOL = ToBool(:StrToInt(:$[1]:):) (ReturnType=IEC_BOOL, ArgType1=IEC_STRING, Inline=Yes)
    STRING_TO_USINT = ToUInt(:StrToInt(:$[1]:),1:) (ReturnType=IEC_USINT, ArgType1=IEC_STRING, Inline=Yes)
    STRING_TO_SINT = ToInt(:StrToInt(:$[1]:),1:) (ReturnType=IEC_SINT, ArgType1=IEC_STRING, Inline=Yes)
    STRING_TO_UINT = ToUInt(:StrToInt(:$[1]:),2:) (ReturnType=IEC_UINT, ArgType1=IEC_STRING, Inline=Yes)
    STRING_TO_INT = ToInt(:StrToInt(:$[1]:),2:) (ReturnType=IEC_INT, ArgType1=IEC_STRING, Inline=Yes)
    STRING_TO_UDINT = ToUInt(:StrToInt(:$[1]:):) (ReturnType=IEC_UDINT, ArgType1=IEC_STRING, Inline=Yes)
    STRING_TO_DINT = ToInt(:StrToInt(:$[1]:):) (ReturnType=IEC_DINT, ArgType1=IEC_STRING, Inline=Yes)
    STRING_TO_REAL = ToFloat(:ToLReal(:$[1]:):) (ReturnType=IEC_REAL, ArgType1=IEC_STRING, Inline=Yes)
    STRING_TO_LREAL = ToLReal(:$[1]:) (ReturnType=IEC_LREAL, ArgType1=IEC_STRING, Inline=Yes)
    LEN = __LEN(:$[1]:) (ReturnType=IEC_INT, ArgType1=IEC_STRING, Inline=Yes)
    LEFT = __LEFT(:$[1], $[2]:) (ReturnType=IEC_STRING, ArgType1=IEC_STRING, ArgType2=IEC_INT, Inline=Yes)
    RIGHT = __RIGHT(:$[1], $[2]:) (ReturnType=IEC_STRING, ArgType1=IEC_STRING, ArgType2=IEC_INT, Inline=Yes)
    MID = __MID(:$[1], $[2], $[3]:) (ReturnType=IEC_STRING, ArgType1=IEC_STRING, ArgType2=IEC_INT, ArgType3=IEC_INT, Inline=Yes)
    CONCAT = __CONCAT(:$[1], $[2]:) (ReturnType=IEC_STRING, ArgType1=IEC_STRING, ArgType2=IEC_STRING, Inline=Yes)
    INSERT = __INSERT(:$[1], $[2], $[3]:) (ReturnType=IEC_STRING, ArgType1=IEC_STRING, ArgType2=IEC_STRING, ArgType3=IEC_INT, Inline=Yes)
    DELETE = __DELETE(:$[1], $[2], $[3]:) (ReturnType=IEC_STRING, ArgType1=IEC_STRING, ArgType2=IEC_INT, ArgType3=IEC_INT, Inline=Yes)
    REPLACE = __REPLACE(:$[1], $[2], $[3], $[4]:) (ReturnType=IEC_STRING, ArgType1=IEC_STRING, ArgType2=IEC_STRING, ArgType3=IEC_INT, ArgType4=IEC_INT, Inline=Yes)
    FIND = __FIND(:$[1], $[2]:) (ReturnType=IEC_INT, ArgType1=IEC_STRING, ArgType2=IEC_STRING, Inline=Yes)
    IP_INST_NUM = IpInstNum(::) (ReturnType=IEC_INT, NumArgs=0)
    IP_OWNER_ID = IpOwnerId(::) (ReturnType=IEC_INT, NumArgs=0)
    PACKET_DATA_ADR = GetIpInt(:6:) (ReturnType=IEC_UDINT, NumArgs=0, Inline=Yes)
    PACKET_COMMAND_ADR = GetIpInt(:7:) (ReturnType=IEC_UDINT, NumArgs=0, Inline=Yes)
  Parameters:
    QUOTED (QuotedName=$R, ValueType=FLOAT, ReturnType=IEC_LREAL)
      ARG (ref=EXPR, DataType=INT, MinValue=0, MaxValue=999)
    QUOTED (QuotedName=$P, ValueType=FLOAT, ReturnType=IEC_LREAL)
      ARG (ref=EXPR, DataType=INT, MinValue=0, MaxValue=999)
    QUOTED (QuotedName=$EXB, ValueType=INT, ReturnType=IEC_SINT)
      ARG (ref=EXPR, DataType=INT, MinValue=0, MaxValue=99)
    QUOTED (QuotedName=$EXW, ValueType=INT, ReturnType=IEC_INT)
      ARG (ref=EXPR, DataType=INT, MinValue=0, MaxValue=99)
    QUOTED (QuotedName=$EXL, ValueType=INT, ReturnType=IEC_DINT)
      ARG (ref=EXPR, DataType=INT, MinValue=0, MaxValue=99)
    QUOTED (QuotedName=$EXF, ValueType=FLOAT, ReturnType=IEC_REAL)
      ARG (ref=EXPR, DataType=INT, MinValue=0, MaxValue=3999)
    QUOTED (QuotedName=$MW, Synchronous=Yes, ValueType=INT, ReturnType=IEC_INT)
      ARG (ref=EXPR, DataType=INT, MinValue=0, MaxValue=99)
    QUOTED (QuotedName=$ML, Synchronous=Yes, ValueType=INT, ReturnType=IEC_DINT)
      ARG (ref=EXPR, DataType=INT, MinValue=0, MaxValue=99)
    QUOTED (QuotedName=$MF, Synchronous=Yes, ValueType=FLOAT, ReturnType=IEC_REAL)
      ARG (ref=EXPR, DataType=INT, MinValue=0, MaxValue=99)
  ParserData (NestedComments=No, DefaultCaseSensitive=Yes, CommentsSpanLines=Yes, ReadWholeFileBeforeParsing=Yes, ExpectMainProgStmts=No, UseFubTemplates=No, LexerType=IEC, RuntimePreventOverflow=No, RoundRealToInt=No, AllowArrayRefWithoutIndex=Yes, DeclareEnumLiteralsAsConstants=No, AllowVariableAutoDereference=Yes, AllowStructMemberAutoDereference=No, AllowPassByRefFnArgAutoReference=No, AllowNamedFnArgs=Yes, AllowUnnamedFnArgs=Yes, AllowFnArgMixedNaming=Yes, AllowFnArgsOutOfSequence=No, AllowBuiltinFnArgsOutOfSequence=Yes, AllowFnArgsOmmitted=Yes, AllowIgnoredFnReturn=Yes, AllowIgnoredExtraSubArgs=No, AllowFnStringInputArgsShort=No, RefuseBuiltinFnUnknownArgName=Yes, AllowBuiltinFnArgCaseSensitive=Yes)
    TKG_OPEN_COMMENT = (*
    TKG_CLOSE_COMMENT = *)
    TKG_IEC_LINE_COMMENT = //
    TKG_TRUE = TRUE:[^\w\d] (IsPattern=Yes)
    TKG_FALSE = FALSE:[^\w\d] (IsPattern=Yes)
    TKG_PRIM_TYPE (IsPattern=Yes)
    TKG_OPEN_BRACKET = (
    TKG_CLOSE_BRACKET = )
    TKG_OPEN_INDEXBRACKET = [
    TKG_CLOSE_INDEXBRACKET = ]
    TKG_COMMA = ,
    TKG_SUBRANGE = ..
    TKG_IEC_BINARY_INTEGER = 2#_[01][01_]+|2#[01][01_]+|2#_[01]|2#[01] (IsPattern=Yes)
    TKG_IEC_OCTAL_INTEGER = 8#_[0-7][0-7_]+|8#[0-7][0-7_]+|8#_[0-7]|8#[0-7] (IsPattern=Yes)
    TKG_IEC_HEX_INTEGER = 16#_[\da-fA-F][\da-fA-F]+|16#[\da-fA-F][\da-fA-F_]+|16#_[\da-fA-F]|16#[\da-fA-F] (IsPattern=Yes)
    TKG_REAL = \d[\d_]*\.[\d_]+[Ee][\+\-]\d[\d_]*|\d[\d_]*\.[\d_]+[Ee]\d[\d_]*|\d[\d_]*\.[\d_]+ (IsPattern=Yes)
    TKG_REAL_EXP = \d[\d_]*[Ee]\d[\d_]*|\d[\d_]*[Ee][\+\-]\d[\d_]* (IsPattern=Yes)
    TKG_INTEGER = \d|\d[\d_]+ (IsPattern=Yes)
    TKG_DOT = .
    TKG_PATHSYNCH_REC_IEC = DO_PATH_SYNCH:[^\w\d] (IsPattern=Yes, EndRuleToken=Yes)
    TKG_PATHSYNCH_END = END_PATH_SYNCH:[^\w\d] (IsPattern=Yes, EndRuleToken=Yes)
    TKG_PATHSYNCH_IPEVAL = IP_EVAL:[^\w\d] (IsPattern=Yes)
    TKG_CYCLIC_PATHSYNCH_BLOCKING_IEC = CYCLIC_PS_BL:[^\w\d] (IsPattern=Yes, EndRuleToken=Yes)
    TKG_CYCLIC_PATHSYNCH_IEC = CYCLIC_PS:[^\w\d] (IsPattern=Yes, EndRuleToken=Yes)
    TKG_CYCLIC_BLOCKING_IEC = CYCLIC_BL:[^\w\d] (IsPattern=Yes, EndRuleToken=Yes)
    TKG_CYCLIC_IEC = CYCLIC:[^\w\d] (IsPattern=Yes, EndRuleToken=Yes)
    TKG_CYCLIC_END_IEC = END_CYCLIC:[^\w\d] (IsPattern=Yes, EndRuleToken=Yes)
    TKG_REFERENCE = REFERENCE:[^\w\d] (FollowedBy=TKG_IEC_TO, IsPattern=Yes)
    TKG_IEC_TO = TO:[^\w\d] (IsPattern=Yes)
    TKG_IEC_DO = DO:[^\w\d] (IsPattern=Yes, EndRuleToken=Yes)
    TKG_FOR_NOFINALDEC = FOR:[^\w\d] (FileXLInvalid=Yes, IsPattern=Yes)
    TKG_FORSTEP = BY:[^\w\d] (FileXLInvalid=Yes, IsPattern=Yes)
    TKG_ENDFOR = END_FOR:[^\w\d] (FileXLInvalid=Yes, IsPattern=Yes, EndRuleToken=Yes)
    TKG_IF = IF:[^\w\d] (IsPattern=Yes)
    TKG_THEN = THEN:[^\w\d] (IsPattern=Yes, EndRuleToken=Yes)
    TKG_BLOCK_ELSEIF = ELSIF:[^\w\d] (IsPattern=Yes)
    TKG_ELSE_AND_DEFAULT = ELSE:[^\w\d] (IsPattern=Yes, EndRuleToken=Yes)
    TKG_BLOCK_ENDIF = END_IF:[^\w\d] (IsPattern=Yes, EndRuleToken=Yes)
    TKG_SWITCH = CASE:[^\w\d] (IsPattern=Yes, FileXLInvalid=Yes)
    TKG_ENDSWITCH_NOBREAK = END_CASE:[^\w\d] (FileXLInvalid=Yes, IsPattern=Yes, EndRuleToken=Yes)
    TKG_WHILE = WHILE:[^\w\d] (FileXLInvalid=Yes, IsPattern=Yes)
    TKG_ENDWHILE = END_WHILE:[^\w\d] (FileXLInvalid=Yes, IsPattern=Yes, EndRuleToken=Yes)
    TKG_DO = REPEAT:[^\w\d] (FileXLInvalid=Yes, IsPattern=Yes, EndRuleToken=Yes)
    TKG_ENDDO_UNTIL = UNTIL:[^\w\d] (FileXLInvalid=Yes, IsPattern=Yes)
    TKG_ENDDO_POSTCOND = END_REPEAT:[^\w\d] (FileXLInvalid=Yes, IsPattern=Yes, EndRuleToken=Yes)
    TKG_BREAK = EXIT:[^\w\d] (FileXLInvalid=Yes, IsPattern=Yes)
    TKG_RETURN = RETURN:[^\w\d] (FileXLInvalid=Yes, IsPattern=Yes)
    TKG_IEC_SEL_FN = SEL:[^\w\d] (FileXLInvalid=Yes, IsPattern=Yes)
    TKG_IEC_MUX_FN = MUX:[^\w\d] (FileXLInvalid=Yes, IsPattern=Yes)
    TKG_TIME_LITERAL = time#\-[dDhHmMsS_\.\d]+|time#[dDhHmMsS_\.\d]+|t#\-[dDhHmMsS_\.\d]+|t#[dDhHmMsS_\.\d]+ (CaseSensitive=no, IsPattern=yes)
    TKG_DATE_AND_TIME_LITERAL = DT#[12]\d\d\d\-[\d\:\-]*|DATE_AND_TIME#[12]\d\d\d\-[\d\:\-]* (CaseSensitive=no, IsPattern=yes)
    TKG_DATE_LITERAL = D#[12]\d\d\d\-[\d\-]*|DATE#[12]\d\d\d\-[\d\-]* (CaseSensitive=no, IsPattern=yes)
    TKG_TIME_OF_DAY_LITERAL = TOD#\d[\d\:\.]*|TIME_OF_DAY#\d[\d\:\.]* (CaseSensitive=no, IsPattern=yes)
    TKG_ASSIGN_EQ = :=
    TKG_OPEN_IP_EXTENSION = {
    TKG_CLOSE_IP_EXTENSION = }
    TKG_IEC_OPEN_TYPE = TYPE:[^\w\d] (IsPattern=Yes)
    TKG_IEC_CLOSE_TYPE = END_TYPE:[^\w\d] (IsPattern=Yes, EndRuleToken=Yes)
    TKG_VAR = VAR:[^\w\d] (IsPattern=Yes)
    TKG_VAR_GLOBAL = VAR_GLOBAL:[^\w\d] (IsPattern=Yes)
    TKG_VAR_INPUT = VAR_INPUT:[^\w\d] (IsPattern=Yes)
    TKG_VAR_OUTPUT = VAR_OUTPUT:[^\w\d] (IsPattern=Yes)
    TKG_VAR_IN_OUT = VAR_IN_OUT:[^\w\d] (IsPattern=Yes)
    TKG_VAR_END = END_VAR:[^\w\d] (IsPattern=Yes, EndRuleToken=Yes)
    TKG_VAR_RETAIN = RETAIN:[^\d\w] (IsPattern=Yes)
    TKG_IP_RETAIN = IP_RETAIN:[^\d\w] (IsPattern=Yes)
    TKG_AT = AT:[^\d\w] (IsPattern=Yes)
    TKG_PLC = PLC:[^\d\w] (IsPattern=Yes)
    TKG_PV_UNDECL = UNRETAIN_VAR:[^\d\w] (IsPattern=Yes)
    TKG_VARSYNCH_IP = IP_SYNCH:[^\d\w] (IsPattern=Yes)
    TKG_VARSYNCH_PATH = PATH_SYNCH:[^\d\w] (IsPattern=Yes)
    TKG_CONSTANT = CONSTANT:[^\d\w] (IsPattern=Yes)
    TKG_VARSCOPE_IP_GLOBAL = IP_GLOBAL:[^\w\d] (IsPattern=Yes)
    TKG_VARSCOPE_SHARED_IP_GLOBAL = SHARED_IP_GLOBAL:[^\w\d] (IsPattern=Yes)
    TKG_VARSCOPE_NC_GLOBAL = NC_GLOBAL:[^\w\d] (IsPattern=Yes)
    TKG_VARSCOPE_PLC_GLOBAL = PLC_GLOBAL:[^\w\d] (IsPattern=Yes)
    TKG_VARSCOPE_IP_LOCAL = LOCAL:[^\w\d] (IsPattern=Yes)
    TKG_IEC_NAMESPACE_SPEC = :: (IsPattern=No)
    TKG_IEC_DATATYPE_SPEC = : (IsPattern=No)
    TKG_IEC_ARRAY = ARRAY:[^\w\d] (IsPattern=Yes)
    TKG_IEC_OF = OF:[^\w\d] (IsPattern=Yes)
    TKG_IEC_DELIM = ; (EndRuleToken=Yes)
    TKG_IEC_OPEN_STRUCT = STRUCT:[^\w\d] (IsPattern=Yes)
    TKG_IEC_CLOSE_STRUCT = END_STRUCT:[^\w\d] (IsPattern=Yes)
    TKG_BITWISE_LP_BINARY_AND = AND:[^\w\d] (IsPattern=Yes)
    TKG_BITWISE_LP_BINARY_OR = OR:[^\w\d] (IsPattern=Yes)
    TKG_BITWISE_LP_BINARY_XOR = XOR:[^\w\d] (IsPattern=Yes)
    TKG_BITWISE_UNARY_COMPLEMENT = NOT:[^\w\d] (IsPattern=Yes)
    TKG_COMP_EXACT_BINARY_GREATER_THAN_OR_EQ = >=
    TKG_COMP_EXACT_BINARY_LESS_THAN_OR_EQ = <=
    TKG_COMP_EXACT_BINARY_EQUAL_TO = =
    TKG_COMP_EXACT_BINARY_NOT_EQUAL_TO = <>
    TKG_COMP_EXACT_BINARY_GREATER_THAN = >
    TKG_COMP_EXACT_BINARY_LESS_THAN = <
    TKG_ARITH_BINARY_PLUS = +
    TKG_ARITH_BINARY_MINUS = -
    TKG_ARITH_BINARY_POWER = **
    TKG_ARITH_BINARY_MULTIPLY = *
    TKG_ARITH_BINARY_DIVIDE = /
    TKG_ARITH_BINARY_MODULO = MOD:[^\w\d] (IsPattern=Yes)
    TKG_PRAGMA = #pragma:[^\w\d] (IsPattern=Yes, FollowedBy=TKG_IDENTIFIER)
    TKG_INCLUDE = #include:[^\w\d] (IsPattern=Yes)
    TKG_PROG_START = PROGRAM:[^\w\d] (IsPattern=Yes, FollowedBy=TKG_PROG_NAME)
    TKG_PROG_NAME = _INIT:[^\w\d]|_CYCLIC:[^\w\d]|_EXIT:[^\w\d]|_MAIN:[^\w\d]|_\d+:[^\w\d] (IsPattern=Yes, EndRuleToken=Yes)
    TKG_PROG_END = END_PROGRAM:[^\w\d] (IsPattern=Yes, EndRuleToken=Yes)
    TKG_SUBPROG_START = FUNCTION:[^\w\d] (IsPattern=Yes)
    TKG_SUBPROG_END = END_FUNCTION:[^\w\d] (IsPattern=Yes, EndRuleToken=Yes)
    TKG_FUB_DECL = FUNCTION_BLOCK:[^\w\d] (IsPattern=Yes)
    TKG_FUB_END = END_FUNCTION_BLOCK:[^\w\d] (IsPattern=Yes, EndRuleToken=Yes)
    TKG_RETURN = RETURN:[^\w\d] (IsPattern=Yes)
    TKG_ACCESS = ACCESS:[^\w\d] (IsPattern=Yes)
    TKG_DEREF_OP = ^
    TKG_ACTION = ACTION:[^\w\d] (IsPattern=Yes)
    TKG_ACTION_END = END_ACTION:[^\w\d] (IsPattern=Yes, EndRuleToken=Yes)
    TKG_IEC_TYPED_VALUE = \w#:[\w\d\+\-]|\w[\w\d]+#:[\w\d\+\-] (IsPattern=Yes)
    TKG_PARAM_PREFIX = $R:[^\w\d]|$P:[^\w\d]|$MW:[^\w\d]|$ML:[^\w\d]|$MF:[^\w\d]|$EXW:[^\w\d]|$EXL:[^\w\d]|$EXF:[^\w\d]|$EXB:[^\w\d] (IsPattern=Yes)
    TKG_IGNORED_IP_EXTENSION = REDUND_CONTEXT|REDUND_UNREPLICABLE|REDUND_OK (IsPattern=Yes)
    TKG_IDENTIFIER = \w|\w[\w\d$]+|$[\w\d$]+ (IsPattern=Yes)
    TKG_INIT_IDENTIFIER = \w|\w[\w\d$]+|$[\w\d$]+ (IsPattern=Yes, Disabled=Yes)
  StringChars (AsciiStringStart=', AsciiStringEnd=', UTF16StringStart=", UTF16StringEnd=")
    EscapeSeq (Search=$N, CaseSensitive=Yes, ReplaceValue=10)
    EscapeSeq (Search=$n, CaseSensitive=Yes, ReplaceValue=10)
    EscapeSeq (Search=$L, CaseSensitive=Yes, ReplaceValue=10)
    EscapeSeq (Search=$l, CaseSensitive=Yes, ReplaceValue=10)
    EscapeSeq (Search=$P, CaseSensitive=Yes, ReplaceValue=12)
    EscapeSeq (Search=$p, CaseSensitive=Yes, ReplaceValue=12)
    EscapeSeq (Search=$R, CaseSensitive=Yes, ReplaceValue=13)
    EscapeSeq (Search=$r, CaseSensitive=Yes, ReplaceValue=13)
    EscapeSeq (Search=$T, CaseSensitive=Yes, ReplaceValue=9)
    EscapeSeq (Search=$t, CaseSensitive=Yes, ReplaceValue=9)
    EscapeSeq (Search=$', CaseSensitive=Yes, ReplaceStr=')
    EscapeSeq (Search=$", CaseSensitive=Yes, ReplaceStr=")
    EscapeSeq (Search=$[\dA-Fa-f]+, IsPattern=Yes, CaseSensitive=Yes, ReplaceEncodingBase=16)
    EscapeSeq (Search=$$, ReplaceStr=$)
    EscapeSeq (Search=$, ReplaceStr=)
```

### Data object Logical/GmcIpConfig/gmciplog (Cnc, version 5.02.1)

#### gmciplog.cnc
```
Root (LangModule=ailgcode, Version=1.0)
  AxesSpec
  PVMacros:
    DR8:
      REF = #next_motion.Data.R8_value
    DI4:
      REF = #next_motion.Data.I4_value
    DU4:
      REF = #next_motion.Data.UI4_value
    DR8_G211:
      SET = %_CNC.TA = ${EXPR};
       if (%_CNC.TA < 0)
         %_CNC.TA = 0;
       endif
        #next_motion.Data.R8_value = ${EXPR};
    Dlp:
      REF = #next_motion.Data.LinMovement.Position
    Dli:
      SET = #next_motion.Data.LinMovement.Idx[0] = ArrayRep(:(:-1:):);
        #next_motion.Data.LinMovement.Idx = ${EXPR};
    Dlm:
      SET = #next_motion.Data.LinMovement.Mode[0] = ArrayRep(:(:-1:):);
        #next_motion.Data.LinMovement.Mode = ${EXPR};
    Dto:
      REF = #next_motion.Data.Trans.Offset
    Dti:
      SET = #next_motion.Data.Trans.AxIdx[0] = ArrayRep(:(:-1:):);
        #next_motion.Data.Trans.AxIdx = ${EXPR};
    Dtm:
      SET = #next_motion.Data.Trans.Mode[0] = ArrayRep(:(:-1:):);
        #next_motion.Data.Trans.Mode = ${EXPR};
    DSPp:
      REF = #next_motion.Data.SplinePoint.Position
    DSPi:
      SET = #next_motion.Data.SplinePoint.AxIdx[0] = ArrayRep(:(:-1:):);
        #next_motion.Data.SplinePoint.AxIdx = ${EXPR};
    DSPm:
      SET = #next_motion.Data.SplinePoint.Mode[0] = ArrayRep(:(:-1:):);
        #next_motion.Data.SplinePoint.Mode = ${EXPR};
    Dcp:
      REF = #next_motion.Data.CircMovement.Parameter
    Dci:
      SET = #next_motion.Data.CircMovement.Idx[0] = ArrayRep(:(:-1:):);
        #next_motion.Data.CircMovement.Idx = ${EXPR};
    Dcm:
      SET = #next_motion.Data.CircMovement.Mode[0] = ArrayRep(:(:-1:):);
        #next_motion.Data.CircMovement.Mode = ${EXPR};
    Dtp:
      REF = #next_motion.Data.ToolAxOrient.Parameter
    Dts:
      REF = #next_motion.Data.ToolAxOrient.Sign
    Daz:
      REF = #next_motion.Data.AbsZeroPtShift.ZpRecIdx
    Das:
      REF = #next_motion.Data.AbsZeroPtShift.SetCS
    Dpt:
      SET = #next_motion.Data.ProgZeroPtShift.Type[0] = ArrayRep(:(:-1:):);
        #next_motion.Data.ProgZeroPtShift.Type = ${EXPR};
    Dpm:
      SET = #next_motion.Data.ProgZeroPtShift.Mode[0] = ArrayRep(:(:-1:):);
        #next_motion.Data.ProgZeroPtShift.Mode = ${EXPR};
    Dpa:
      REF = #next_motion.Data.ProgZeroPtShift.AxShift
    Dovpathdef:
      REF = #next_motion.Data.OptMotPar.path_definition
    Dovpathdefd:
      REF = #next_motion.Data.OptMotPar.path_definition_def
    Dorpar:
      REF = #next_motion.Data.OptMotPar.robot_par
    Dorpard:
      REF = #next_motion.Data.OptMotPar.robot_par_def
    Dolim:
      REF = #next_motion.Data.OptMotPar.limits_idx
    Dolimd:
      REF = #next_motion.Data.OptMotPar.limits_idx_def
    Dolimfac:
      REF = #next_motion.Data.OptMotPar.limits_factor
    Dolimfacd:
      REF = #next_motion.Data.OptMotPar.limits_factor_def
    Dfdx:
      REF = #next_motion.Data.FullTrfTool.Dx
    Dfdy:
      REF = #next_motion.Data.FullTrfTool.Dy
    Dfdz:
      REF = #next_motion.Data.FullTrfTool.Dz
    Dfph:
      REF = #next_motion.Data.FullTrfTool.Phi
    Dft:
      REF = #next_motion.Data.FullTrfTool.Theta
    Dfps:
      REF = #next_motion.Data.FullTrfTool.Psi
    DPLDli:
      REF = #next_motion.Data.PosLatchDistance.LatchIdx
    DPLDts:
      REF = #next_motion.Data.PosLatchDistance.TriggSource
    DPLDe:
      REF = #next_motion.Data.PosLatchDistance.Edge
    DPLDti:
      REF = #next_motion.Data.PosLatchDistance.HwTrigIdx
    DPLDd:
      REF = #next_motion.Data.PosLatchDistance.Distance
    DPLli:
      REF = #next_motion.Data.PosLatch.LatchIdx
    DPLts:
      REF = #next_motion.Data.PosLatch.TriggSource
    DPLe:
      REF = #next_motion.Data.PosLatch.Edge
    DPLti:
      REF = #next_motion.Data.PosLatch.HwTrigIdx
    DPLtr:
      REF = #next_motion.Data.PosLatchGmc.Trigger
    DPLlp:
      REF = #next_motion.Data.PosLatchGmc.pLatchPos
    DPLcs:
      REF = #next_motion.Data.PosLatchGmc.CoordSystem
    DPLrp:
      REF = #next_motion.Data.PosLatchGmc.ResidualPath
    Drma:
      REF = #next_motion.Data.R_DependFeed.MaxRadius
    Drmi:
      REF = #next_motion.Data.R_DependFeed.MinRadius
    Drr:
      REF = #next_motion.Data.R_DependFeed.Rate
    Dsvp:
      SET = #next_motion.Data.Set_v_jump.programmed[0] = ArrayRep(:(:ncOFF:):);
        #next_motion.Data.Set_v_jump.programmed = ${EXPR};
    Dsvv:
      REF = #next_motion.Data.Set_v_jump.value
    Dsap:
      SET = #next_motion.Data.Set_a_jump.programmed[0] = ArrayRep(:(:ncOFF:):);
        #next_motion.Data.Set_a_jump.programmed = ${EXPR};
    Dsav:
      REF = #next_motion.Data.Set_a_jump.value
    Dsep:
      SET = #next_motion.Data.SetAxLimit.programmed[0] = ArrayRep(:(:ncOFF:):);
        #next_motion.Data.SetAxLimit.programmed = ${EXPR};
    Dser:
      REF = #next_motion.Data.SetAxLimit.RecordIdx
    Dcad:
      REF = #next_motion.Data.CamWrapping.Diameter
    Dcap:
      REF = #next_motion.Data.CamWrapping.ParameterP1
    Dsu:
      REF = #next_motion.Data.SetPathAccDec.UnitType
    Dsv108:
      SET = #next_motion.Data.SetPathAccDec.value = ${EXPR};
        if (#next_motion.Data.SetPathAccDec.UnitType == 1)
          %_CNC.lim_path_acc_p = ${EXPR} / 100.0 * %_CNC.lim_path_acc_p_ini;
        else
          %_CNC.lim_path_acc_p = ${EXPR};
        endif
    Dsv109:
      SET = #next_motion.Data.SetPathAccDec.value = ${EXPR};
        if (#next_motion.Data.SetPathAccDec.UnitType == 1)
          %_CNC.lim_path_acc_n = ${EXPR} / 100.0 * %_CNC.lim_path_acc_n_ini;
        else
          %_CNC.lim_path_acc_n = ${EXPR};
        endif
    Dsv110:
      SET = #next_motion.Data.SetPathAccDec.value = ${EXPR};
        if (#next_motion.Data.SetPathAccDec.UnitType == 1)
          %_CNC.lim_path_acc_p = ${EXPR} / 100.0 * %_CNC.lim_path_acc_p_ini;
          %_CNC.lim_path_acc_n = ${EXPR} / 100.0 * %_CNC.lim_path_acc_n_ini;
        else
          %_CNC.lim_path_acc_p = ${EXPR};
          %_CNC.lim_path_acc_n = ${EXPR};
        endif
    Daxlv:
      REF = #next_motion.Data.AxisLimit.Value
    Daxla:
      REF = #next_motion.Data.AxisLimit.Axis
    Daxlu:
      REF = #next_motion.Data.AxisLimit.UnitType
    Dsma:
      REF = #next_motion.Data.SetTransSpeed.MaxAngle
    Dsmi:
      REF = #next_motion.Data.SetTransSpeed.MinAngle
    Dsr:
      REF = #next_motion.Data.SetTransSpeed.RedFactor
    Dbrp:
      REF = #next_motion.Data.BezierSpline.RadiusProgrammed
    Dbr:
      REF = #next_motion.Data.BezierSpline.Radius
    Dbvp:
      REF = #next_motion.Data.BezierSpline.VeProgrammed
    Dbv:
      REF = #next_motion.Data.BezierSpline.Ve
    Dbl:
      REF = #next_motion.Data.BezierSpline.LinProgrammed
    Dbsf:
      REF = #next_motion.Data.BezierSpline.scalingFactor
    Dbsfd:
      REF = #next_motion.Data.BezierSpline.scalingFactor_def
    Dao:
      REF = #next_motion.Data.AutomTangentialAx.Offset
    Daa:
      REF = #next_motion.Data.AutomTangentialAx.AxIdx
    DAMa:
      REF = #next_motion.Data.AxisMapping.AxIdx
    DAMf:
      REF = #next_motion.Data.AxisMapping.factor
    DAMp:
      REF = #next_motion.Data.AxisMapping.ParameterP1
    DSPEid:
      REF = #next_motion.Data.SignalPathEnd.SignalId
    DSPEt:
      REF = #next_motion.Data.SignalPathEnd.Time
    DSPEst:
      REF = #next_motion.Data.SignalPathEnd.SignalType
    DSPEsi:
      REF = #next_motion.Data.SignalPathEnd.SignalIdx
    DSPEsd:
      REF = #next_motion.Data.SignalPathEnd.SourceData
    DSPEd:
      REF = #next_motion.Data.SignalPathEnd.DataLength
    DSPEp:
      SET = #next_motion.Data.SignalPathEnd.pDestination = \#sys_vars.EXF[0];
    DSPEDid:
      REF = #next_motion.Data.SignalPathEndDist.SignalId
    DSPEDd:
      REF = #next_motion.Data.SignalPathEndDist.Distance
    DSPEDst:
      REF = #next_motion.Data.SignalPathEndDist.SignalType
    DSPEDsi:
      REF = #next_motion.Data.SignalPathEndDist.SignalIdx
    DSPEDsd:
      REF = #next_motion.Data.SignalPathEndDist.SourceData
    DSPEDdl:
      REF = #next_motion.Data.SignalPathEndDist.DataLength
    DSPEDp:
      SET = #next_motion.Data.SignalPathEndDist.pDestination = \#sys_vars.EXF[0];
    DSPo:
      REF = #next_motion.Data.SignalPredict.Override
    DSPop:
      REF = #next_motion.Data.SignalPredict.OvrProgrammed
    DSPsi:
      REF = #next_motion.Data.SignalPredict.SignalIdx
    DSPsp:
      REF = #next_motion.Data.SignalPredict.StopProgrammed
    DWCx1:
      REF = #next_motion.Data.WS_Ctrl.x1
    DWCz1:
      REF = #next_motion.Data.WS_Ctrl.z1
    DWCy1:
      REF = #next_motion.Data.WS_Ctrl.y1
    DWCx2:
      REF = #next_motion.Data.WS_Ctrl.x2
    DWCz2:
      REF = #next_motion.Data.WS_Ctrl.y2
    DWCy2:
      REF = #next_motion.Data.WS_Ctrl.z2
    DWCi:
      REF = #next_motion.Data.WS_Ctrl.index
    DWCc:
      REF = #next_motion.Data.WS_Ctrl.coord
    DWCpl:
      REF = #next_motion.Data.WS_Ctrl.pplane
    DWCo:
      REF = #next_motion.Data.WS_Ctrl.orient
    DWCs:
      REF = #next_motion.Data.WS_Ctrl.shape
    DWCca:
      REF = #next_motion.Data.WS_Ctrl.clear_all
    DWCp1:
      REF = #next_motion.Data.WS_Ctrl.point1
    DWCp2:
      REF = #next_motion.Data.WS_Ctrl.point2
    DWCen:
      REF = #next_motion.Data.WS_Ctrl.enable
    DWCa:
      SET = #next_motion.Data.WS_Ctrl.arm_diameter[0] = ArrayRep(:(:ncOFF:):);
        #next_motion.Data.WS_Ctrl.arm_diameter = ${EXPR};
    DTDRt:
      REF = #next_motion.Data.ToolDataRecord.ToolIdx
    Sz:
      REF = #sys_vars.ZP
    DSSi:
      REF = #next_motion.Data.SpindleSpeed.Idx
    DSSs:
      REF = #next_motion.Data.SpindleSpeed.speed
    DCSSt:
      REF = #next_motion.Data.C2_SplineStart.BCType
    DCSSv:
      REF = #next_motion.Data.C2_SplineStart.BCValue
    DCSSp:
      SET = #next_motion.Data.C2_SplineStart.BCProgrammed[0] = ArrayRep(:(:ncOFF:):);
        #next_motion.Data.C2_SplineStart.BCProgrammed = ${EXPR};
    DCSSsp:
      REF = #next_motion.Data.C2_SplineStart.SegmentParameter
    DCSSst:
      REF = #next_motion.Data.C2_SplineStart.SegmentType
    DCSEt:
      REF = #next_motion.Data.C2_SplineEnd.BCType
    DCSEv:
      REF = #next_motion.Data.C2_SplineEnd.BCValue
    DCSEp:
      SET = #next_motion.Data.C2_SplineEnd.BCProgrammed[0] = ArrayRep(:(:ncOFF:):);
        #next_motion.Data.C2_SplineEnd.BCProgrammed = ${EXPR};
    DFd:
      REF = #next_motion.Data.Frame.Data
    DFcs:
      REF = #next_motion.Data.Frame.SetCS
    DSVs:
      REF = #next_motion.Data.SystemVariable.SysVarIdx
    DSVa:
      REF = #next_motion.Data.SystemVariable.AxIdx
    DSVd:
      REF = #next_motion.Data.SystemVariable.Data.R8_value
    DABNf:
      REF = #next_motion.Data.AutoBlockNumber.offset
    DABNo:
      REF = #next_motion.Data.AutoBlockNumber.factor
    DCSSPs:
      REF = #next_motion.Data.ConstantSurfaceSpeed.Speed
    DCSSPp:
      REF = #next_motion.Data.ConstantSurfaceSpeed.Programmed
    MXFPx:
      REF = #next_motion.Data.MXFrame.Pos.x
    MXFPy:
      REF = #next_motion.Data.MXFrame.Pos.y
    MXFPz:
      REF = #next_motion.Data.MXFrame.Pos.z
    MXFOt:
      REF = #next_motion.Data.MXFrame.Orient.Type
    MXFOa:
      REF = #next_motion.Data.MXFrame.Orient.Angle
    MXFEPx:
      REF = #next_motion.Data.MXFrameEx.Frame.Pos.x
    MXFEPy:
      REF = #next_motion.Data.MXFrameEx.Frame.Pos.y
    MXFEPz:
      REF = #next_motion.Data.MXFrameEx.Frame.Pos.z
    MXFEOt:
      REF = #next_motion.Data.MXFrameEx.Frame.Orient.Type
    MXFEOa:
      REF = #next_motion.Data.MXFrameEx.Frame.Orient.Angle
    MXFECs:
      REF = #next_motion.Data.MXFrameEx.SetCS
    MXFEAd:
      REF = #next_motion.Data.MXFrameEx.Additive
    MXTFPx:
      REF = #next_motion.Data.MXTool.Frame.Pos.x
    MXTFPy:
      REF = #next_motion.Data.MXTool.Frame.Pos.y
    MXTFPz:
      REF = #next_motion.Data.MXTool.Frame.Pos.z
    MXTFOt:
      REF = #next_motion.Data.MXTool.Frame.Orient.Type
    MXTFOa:
      REF = #next_motion.Data.MXTool.Frame.Orient.Angle
    MXTr:
      REF = #next_motion.Data.MXTool.Radius
    MXTi:
      REF = #next_motion.Data.MXTool.Index
    MXPPx:
      REF = #next_motion.Data.MXPoint.Pos.x
    MXPPy:
      REF = #next_motion.Data.MXPoint.Pos.y
    MXPPz:
      REF = #next_motion.Data.MXPoint.Pos.z
    MXPOt:
      REF = #next_motion.Data.MXPoint.Orient.Type
    MXPOa:
      REF = #next_motion.Data.MXPoint.Orient.Angle
    MXPCm:
      REF = #next_motion.Data.MXPoint.Cfg.Mode
    MXPr:
      REF = #next_motion.Data.MXPoint.RotAxis
    MXPa:
      REF = #next_motion.Data.MXPoint.AuxAxis
    MXPhTr:
      REF = #next_motion.Data.MXPathDesc.Trans.Radius
    MXPhTt:
      REF = #next_motion.Data.MXPathDesc.Trans.Type
    MXDa:
      REF = #next_motion.Data.MXDynamicDesc.Accel
    MXDd:
      REF = #next_motion.Data.MXDynamicDesc.Decel
    MXDOe:
      REF = #next_motion.Data.MXDynamicDesc.Optmot.Enable
    MXDOv:
      REF = #next_motion.Data.MXDynamicDesc.Optmot.VelPathDef
    MXDOr:
      REF = #next_motion.Data.MXDynamicDesc.Optmot.RobotPar
    MXDOl:
      REF = #next_motion.Data.MXDynamicDesc.Optmot.Limits
    MXVv:
      REF = #next_motion.Data.MXVelocity.v
    MXVm:
      REF = #next_motion.Data.MXVelocity.Mode
    MXAj:
      REF = #next_motion.Data.MXAxisTarget.JointAxis
    MXAa:
      REF = #next_motion.Data.MXAxisTarget.AuxAxis
    MXAb:
      REF = #next_motion.Data.MXAxisTarget.BaseAxis
    MXJ:
      REF = #next_motion.Data.MXJointAxis
    MXAto:
      REF = #next_motion.Data.MXAutoTang.Offset
    MXCDCas:
      REF = #next_motion.Data.MXCDC.ArcTransSpd
    MXCDCsm:
      REF = #next_motion.Data.MXCDC.SpdMode
    MXCDCcv:
      REF = #next_motion.Data.MXCDC.ContourViolation
    MXCDCtm:
      REF = #next_motion.Data.MXCDC.TransMode
    MXCDCem:
      REF = #next_motion.Data.MXCDC.EntryMode
    MXCDCal:
      REF = #next_motion.Data.MXCDC.AcrToLine
    THCp:
      REF = #next_motion.Data.ThreadCut.Position
    THCi:
      SET = #next_motion.Data.ThreadCut.Idx[0] = ArrayRep(:(:-1:):);
        #next_motion.Data.ThreadCut.Idx = ${EXPR};
    THCm:
      SET = #next_motion.Data.ThreadCut.Mode[0] = ArrayRep(:(:-1:):);
        #next_motion.Data.ThreadCut.Mode = ${EXPR};
    THCld:
      REF = #next_motion.Data.ThreadCut.LeadDirection
    THCl:
      REF = #next_motion.Data.ThreadCut.Lead
    THCo:
      REF = #next_motion.Data.ThreadCut.Offset
    ACVc:
      REF = #next_motion.Data.AxisCtrlVelocity.Command
    ACVi:
      REF = #next_motion.Data.AxisCtrlVelocity.Idx
    ACSs:
      REF = #next_motion.Data.AxisCtrlSpeed.Speed
    ACSi:
      REF = #next_motion.Data.AxisCtrlSpeed.Idx
    ACPp:
      REF = #next_motion.Data.AxisCtrlPosition.Position
    ACPd:
      REF = #next_motion.Data.AxisCtrlPosition.PositionDefined
    ACPi:
      REF = #next_motion.Data.AxisCtrlPosition.Idx
    ACPm:
      REF = #next_motion.Data.AxisCtrlPosition.Mode
    CHFm:
      REF = #next_motion.Data.Chamfer.Mode
    CHFv:
      REF = #next_motion.Data.Chamfer.Value
    PAFv:
      REF = #next_motion.Data.PathFeed.Value
    PAFi:
      REF = #next_motion.Data.PathFeed.Id
    GENd:
      REF = #next_motion.Data.GenericData.Data
    SGALda:
      REF = #next_motion.Data.SetGmcAxisLimit.DestinationAxis
    SGALdp:
      REF = #next_motion.Data.SetGmcAxisLimit.DestinationPath
    SGALsa:
      REF = #next_motion.Data.SetGmcAxisLimit.SourceAxis
    SGALsp:
      REF = #next_motion.Data.SetGmcAxisLimit.SourcePath
    SGALn:
      SET = BlockCpy(:\#next_motion.Data.SetGmcAxisLimit.SourceLimitSetName, ${EXPR}:);
    CMPmd:
      REF = #next_motion.Data.Compressor.MaxCartesianDeviation
    CMPmnd:
      REF = #next_motion.Data.Compressor.MaxNonCartesianDeviation
    CMPmt:
      REF = #next_motion.Data.Compressor.MaxCartesianTransitionAngle
    CMPml:
      REF = #next_motion.Data.Compressor.MaxCartesianLength
    CMPmnt:
      REF = #next_motion.Data.Compressor.MaxNonCartesianTransitionAngle
    PR8v:
      REF = #next_motion.Data.R8_param.Value
    PR8i:
      REF = #next_motion.Data.R8_param.Id
    STPi:
      REF = #next_motion.Data.ToolPar.Id
    STPR8:
      REF = #next_motion.Data.ToolPar.R8_value
    STPI4:
      REF = #next_motion.Data.ToolPar.I4_value
    GFof:
      REF = #next_motion.Data.GmcFrame.Offset
    GFmo:
      SET = #next_motion.Data.GmcFrame.Mode[0] = ArrayRep(:(:-1:):);
        #next_motion.Data.GmcFrame.Mode = ${EXPR};
    GFai:
      SET = #next_motion.Data.GmcFrame.AxIdx[0] = ArrayRep(:(:-1:):);
        #next_motion.Data.GmcFrame.AxIdx = ${EXPR};
    GFor:
      REF = #next_motion.Data.GmcFrame.Orientation
    GFori:
      SET = #next_motion.Data.GmcFrame.OrientationIdx[0] = ArrayRep(:(:-1:):);
        #next_motion.Data.GmcFrame.OrientationIdx = ${EXPR};
    GFort:
      REF = #next_motion.Data.GmcFrame.OrientationType
    GFsc:
      REF = #next_motion.Data.GmcFrame.SetCS
    GFtfc:
      REF = #next_motion.Data.GmcFrame.TCPFromCS
    GFttc:
      REF = #next_motion.Data.GmcFrame.TCPToCS
    GFcc:
      REF = #next_motion.Data.GmcFrame.ClearCS
    GFne:
      REF = #next_motion.Data.GmcFrame.Negative
    GFut:
      REF = #next_motion.Data.GmcFrame.UseTCP
  Constants:
    PathBusy = BUSY (type=STRING)
    PathStatus = STATUS (type=STRING)
    PathErrLevel = ERRLEV (type=STRING)
  BuiltInProcs:
    SendCommand = SendCommand(:$[1]:); (MinArgs=1, MaxArgs=1, Inline=Yes)
    DispatchAndWait = DispatchAndWait(:$[1]:); (MinArgs=1, MaxArgs=1, Inline=Yes)
    WaitForCommand = WaitForCommand(:$[1]:); (MinArgs=1, MaxArgs=1, Inline=Yes)
  Preprocess:
    MP_PJN (Search=MP22000 , Replace=PJN )
    MP_PJB (Search=MP22100 , Replace=PJB )
  GCodes:
    G_DELAY (GNum=0, Alias=@, AliasIsPattern=Yes, Inline=Yes)
      Arg (DataType=FLOAT, ref=tickdelay)
    G_PJN (GNum=22000, Alias=PJN, Group=220)
      Arg PathBusy (DataType=FLOAT, ref=busy_count)
      Arg PathStatus (DataType=FLOAT, ref=final_status)
      Arg PathErrLevel (DataType=FLOAT, ref=error_level)
    G_PJB (GNum=22100, Alias=PJB, Group=220)
      Arg PathBusy (DataType=FLOAT, ref=busy_count)
      Arg PathStatus (DataType=FLOAT, ref=final_status)
      Arg PathErrLevel (DataType=FLOAT, ref=error_level)
  MCodes:
    M_DEFAULT (IsDefault=Yes, MinValue=0, MaxValue=999999)
      ARG (ref=VALUE, DataType=FLOAT, RequireLiteral=Yes)
    M10003 = 10003 (Inline=Yes)
      ARG (ref=VALUE, DataType=FLOAT, RequireLiteral=Yes)
    M1000000 = 1000000 (Alias=;, AliasIsPattern=Yes, Inline=Yes, IgnoreIfGroups=220)
      ARG (ref=VALUE, DataType=FLOAT, RequireLiteral=Yes)
  ParserData (NestedComments=No, DefaultCaseSensitive=Yes, CommentsSpanLines=No, ReadWholeFileBeforeParsing=No, ExpectMainProgStmts=Yes, UseFubTemplates=No)
    TKG_END_OF_LINE = \n (IsPattern=No)
    TKG_OPEN_COMMENT = #
    TKG_NC_BLOCK_PREFIX = N:[\s\d] (IsPattern=Yes)
    TKG_OPEN_LISTBRACKET = (
    TKG_CLOSE_LISTBRACKET = )
    TKG_COMMA = ,
    TKG_NUMBER = \d+\.\d+|\d+\.|\.\d+ (IsPattern=Yes)
    TKG_INTEGER = \d+ (IsPattern=Yes)
    TKG_NUMBER_EXP = e:[\s\d\+\-\.] (IsPattern=Yes)
    TKG_ASSIGN_EQ = =
    TKG_ARITH_BINARY_MINUS = -
    TKG_M_CODE_PREFIX = MP:\d (IsPattern=Yes)
  StringChars (AsciiStringStart=")
    EscapeSeq (Search=$N, CaseSensitive=No, ReplaceValue=10)
    EscapeSeq (Search=$L, CaseSensitive=Yes, ReplaceValue=10)
    EscapeSeq (Search=$Q, CaseSensitive=No, ReplaceStr=")
    EscapeSeq (Search=$[\dA-F]+, IsPattern=Yes, CaseSensitive=No, ReplaceEncodingBase=16)
    EscapeSeq (Search=$$, ReplaceStr=$)
    EscapeSeq (Search=$, ReplaceStr=)
```

### Data object Logical/GmcIpConfig/gmcipesm (Cnc, version 5.02.1)
